      | #           return OBJECT_MAP[i]
      | #       end
      | #       i = i + 1
      | #   end
      | #   return OBJ_DEFAULT  # Return default pattern if not found
      | # end
      | 
      | def find_object_by_objectname(objectname):
      |     local i = 0
      |     #log_info("Trying to find object by color:", to_str(objectname))
      |     while (i < OBJECT_MAP.length()):
      |         if (OBJECT_MAP[i].obj_name == objectname):
      |             log_info("Object Model found: [" + to_str(OBJECT_MAP[i].description) + "]")
      |             return OBJECT_MAP[i]
      |         end
      |         i = i + 1
      |     end
      |     log_warning("no Object Model found for objectname:[" + to_str(objectname) + "]")
      |     return create_object()
      | end
      | 
      | def find_smallest_object():
      |     local i = 0
      |     local min_size = OBJECT_MAP[0].height
      |     #log_info("Trying to find object by color:", to_str(objectname))
      |     while (i < OBJECT_MAP.length()):
      |         if (OBJECT_MAP[i].height <= min_size and OBJECT_MAP[i].height != 0):
      |             log_info("smaller object found: [" + to_str(OBJECT_MAP[i].description) + "]")
      |             min_size = OBJECT_MAP[i].height
      |         end
      |         i = i + 1
      |     end
      |     return min_size
      | end
      | 
      | def find_gripper_config_by_objectname(objectname):
      | local i = 0
      | while (i < GRIPPER_CONFIG_MAP.length()):
      |     #log_info("gripper config:",to_str(GRIPPER_CONFIG_MAP[i]))
      |     if (GRIPPER_CONFIG_MAP[i].object == objectname):
      |         log_info("found gripper parameters [" + to_str(GRIPPER_CONFIG_MAP[i]) + "]")
      |         return GRIPPER_CONFIG_MAP[i]
      |     end
      |     i = i + 1
      | end
      | 
      | log_warning("no gripper parameters found for object type: " + to_str(objectname))
      | return create_gripper_config()
      | end
      | # Function to find a landmark by item
      | def find_landmark_by_id(lm_id):
      |     local i = 0
      |     while i < LANDMARK_MAP.length():
      |         if LANDMARK_MAP[i].lm_id == lm_id:
      |             log_info("found landmark with id(" + to_str(lm_id) + "): [" + to_str(LANDMARK_MAP[i].description) + "]")
      |             return LANDMARK_MAP[i]
      |         end
      |         i = i + 1
      |     end
      |     log_warning("landmark not found for lm_id [" + to_str(lm_id) + "]")
      |     return create_landmark()
      | end
      | # Function to find a landmark by item
      | def find_landmark_by_capture_pos(capture_pos):
      |     local i = 0
      |     while i < LANDMARK_MAP.length():
      |         if LANDMARK_MAP[i].capture_pos == capture_pos:
      |             log_info("found landmark by capture_pos [" + to_str(LANDMARK_MAP[i].description) + "]")
      |             return LANDMARK_MAP[i]
      |         end
      |         i = i + 1
      |     end
      |     log_warning("Landmark not found for capture_pos: [" + to_str(capture_pos) + "]")
      |     return create_landmark()
      | end
      | 
      | def update_landmark_by_capture_pos(capture_pos, lm_pos):
      |     local i = 0
      |     while i < LANDMARK_MAP.length():
      |         if LANDMARK_MAP[i].capture_pos == capture_pos:
      |             log_info("updated landmark from [" + to_str(LANDMARK_MAP[i].description) + "]")
      |             LANDMARK_MAP[i].actual_frame = lm_pos
      |             return True
      |         end
      |         i = i + 1
      |     end
      |     log_warning("Landmark not found for capture_pos: [" + to_str(capture_pos) + "]")
      |     return False
      | end
      | 
      | def update_landmark_by_id(lm_id,lm_pos):
      |     local i = 0
      |     while i < LANDMARK_MAP.length():
      |         if LANDMARK_MAP[i].lm_id == lm_id:
      |             log_info("updated landmark.actual_frame from [" + to_str(LANDMARK_MAP[i].description + "]"))
      |             LANDMARK_MAP[i].actual_frame = lm_pos
      |             return True
      |         end
      |         i = i + 1
      |     end
      |     log_warning("Landmark not found for lm_id " + to_str(lm_id))
      |     return False
      | end
      | 
      | def find_vision_config_by_frame(frame):
      |     local i = 0
      |     while i < VISION_CONFIG_MAP.length():
      |         if VISION_CONFIG_MAP[i].capture_pos == frame:
      |             log_info("Vision Config found: [" + to_str(VISION_CONFIG_MAP[i].description) + "]")
      |             return VISION_CONFIG_MAP[i]
      |         end
      |         i = i + 1
      |     end
      |     log_info("Vision Config not found for frame: " + to_str(frame))
      |     return create_vision_config()
      | end
      | 
      | def find_vision_config_by_itemid(id):
      |     local i = 0
      |     while i < VISION_CONFIG_MAP.length():
      |         if VISION_CONFIG_MAP[i].item_id == id:
      |             log_info("Vision Config found: [" + to_str(VISION_CONFIG_MAP[i].description) + "]")
      |             return VISION_CONFIG_MAP[i]
      |         end
      |         i = i + 1
      |     end
      |     log_info("Vision Config not found for item: " + to_str(id))
      |     return create_vision_config()
      | end
      | 
      | def find_inspect_config_by_itemid(id):
      |     local i = 0
      |     while i < INSPECT_CONFIG_MAP.length():
      |         if INSPECT_CONFIG_MAP[i].item_id == id:
      |             log_info("Inspect Config found: [" + to_str(INSPECT_CONFIG_MAP[i].description) + "]")
      |             return INSPECT_CONFIG_MAP[i]
      |         end
      |         i = i + 1
      |     end
      |     log_info("Inspect Config not found for item: " + to_str(id))
      |     return create_inspect_config()
      | end
    Script file /programs/04 Scripts/SCRIPT Device Robotiq Greifer v0.2.script
      | # ############ SCRIPT Device Robotiq Greifer ###############
      | # **********************************************************
      | # Customer          :   URG
      | # Product Name      :   uLabMobile
      | # **********************************************************
      | # Controller/Robot  :   UR5e
      | # Software          :   5.17
      | # Dependencies      :   Logs Script, Robotiq Gripper and Gripper Datastructure for args (Factory Script), URCAP Robotiq
      | # **********************************************************
      | # Author            :   D.Kreugel, P.Köhnke
      | # Copyright (c)     :   United Robotics Group Health and Food GmbH
      | #                       An der Riede 2
      | #                       28816 Stuhr
      | #                       Germany
      | # *********************************************************
      | # Description       :   Gripper Robotiq Device Interface for Robotiq E-Hand Gripper
      | # Version           :   0.2
      | # Created           :   18.07.2024
      | # Updated           :
      | # *********************************************************
      | # Modifications     :
      | #
      | # Date              :
      | # Name              :
      | # Reason            :
      | # *********************************************************
      | # TODO              :   documentation
      | 
      | # RobotiQ Gripper
      | ROBOTIQ_GRP_CLOSE = 0
      | ROBOTIQ_GRP_OPEN = 40
      | 
      | # #############FORCEMODE###############
      | ROBOTIQ_GRP_FORCE = struct(FULL=100, HALF=50, LOW=25, NONE=0)
      | 
      | # #############SPEED###################
      | ROBOTIQ_GRP_SPEED = struct(FAST=100, MEDIUM=50, SLOW=20)
      | 
      | # ############VALIDATION###############
      | ROBOTIQ_GRP_VALIDATION = struct(ON=1, OFF=0, SKIP=-1)
      | 
      | # struct(prepick=0, pick=0, place=0, force=0, speed=0, validation=0, object_type=0, description="default")
      | def gripper_robotiq_activate():
      |     return rq_activate_and_wait()
      | end
      | 
      | def gripper_robotiq_reset_and_activate():
      |     return rq_reset_and_activate()
      |     #return rq_reset()
      | end
      | 
      | def gripper_robotiq_is_activated():
      |     return rq_is_gripper_activated()
      | end
      | 
      | def gripper_robotiq_get_current_pos_mm():
      |     return rq_current_pos_mm()
      | end
      | # Function to check if the RobotiQ gripper has an object
      | def gripper_robotiq_has_object():
      |     result = rq_is_object_detected()
      |     if result == False:
      |         log_error("No object detected by the gripper")
      |     end
      |     return result
      | end
      | 
      | def gripper_robotiq_move_to_mm(mm):
      |     if(gripper_robotiq_is_activated() == False):
      |         gripper_robotiq_activate()
      |     end
      |     return rq_move_and_wait_mm(mm)
      | end
      | 
      | def gripper_robotiq_close():
      |     if(gripper_robotiq_is_activated() == False):
      |         gripper_robotiq_activate()
      |     end
      |     return rq_close_and_wait()
      | end
      | 
      | def gripper_robotiq_open():
      |     if(gripper_robotiq_is_activated() == False):
      |         gripper_robotiq_activate()
      |     end
      |     return rq_open_and_wait()
      | end
      | 
      | def gripper_robotiq_set_force(force):
      |     return rq_set_force_norm(force)
      | end
      | 
      | def gripper_robotiq_set_speed(velocity):
      |     return rq_set_speed_norm(velocity)
      | end
      | # Function to initialize the RobotiQ gripper
      | # args = struct(obj_type = object.obj_type, force = force, speed = speed, validation = validation, width = (prepick=2, pick=0, place=2))
      | def gripper_robotiq_init(args):
      |     log_info("args:"+to_str(args))
      |     gripper_robotiq_set_force(args.force)
      |     gripper_robotiq_set_speed(args.speed)
      |     if(gripper_robotiq_is_activated() == False):
      |         gripper_robotiq_activate()
      |     end
      |     log_info("Robotiq Gripper Initialized with arguments:" + to_str(args))
      |     return True
      | end
      | # Function to prepare the RobotiQ gripper for picking
      | # args = struct(obj_type = object.obj_type, force = force, speed = speed, validation = validation, width = (prepick=2, pick=0, place=2))
      | def gripper_robotiq_prepick(args):
      |     gripper_robotiq_init(args)
      | 
      |     if(args.width.prepick <= ROBOTIQ_GRP_CLOSE):
      |         rq_close_and_wait()
      |     elif(args.width.prepick >= ROBOTIQ_GRP_OPEN):
      |         rq_open_and_wait()
      |     else:
      |         rq_move_and_wait_mm(args.width.prepick)
      |     end
      | 
      |     log_info("Robotiq Gripper prepick with arguments:" + to_str(args))
      |     return True
      | end
      | 
      | # Function to place an object using the RobotiQ gripper
      | # args = struct(obj_type = object.obj_type, force = force, speed = speed, validation = validation, width = (prepick=2, pick=0, place=2))
      | def gripper_robotiq_place(args):
      |     gripper_robotiq_init(args)
      | 
      |     if(args.width.place <= ROBOTIQ_GRP_CLOSE):
      |         rq_close_and_wait()
      |     elif(args.width.place >= ROBOTIQ_GRP_OPEN):
      |         rq_open_and_wait()
      |     else:
      |         rq_move_and_wait_mm(args.width.place)
      |     end
      | 
      |     log_info("Gripper Place with arguments:"+ to_str(args))
      |     return True
      | end
      | 
      | # Function to pick an object using the RobotiQ gripper
      | # args = struct(obj_type = object.obj_type, force = force, speed = speed, validation = validation, width = (prepick=2, pick=0, place=2))
      | def gripper_robotiq_pick(args):
      |     gripper_robotiq_init(args)
      | 
      |     if(args.width.pick <= ROBOTIQ_GRP_CLOSE):
      |         rq_close_and_wait()
      |     elif(args.width.pick >= ROBOTIQ_GRP_OPEN):
      |         rq_open_and_wait()
      |     else:
      |         rq_move_and_wait_mm(args.width.pick)
      |     end
      | 
      |     log_info("Gripper Pick with arguments:" + to_str(args))
      | 
      |     if args.validation == ROBOTIQ_GRP_VALIDATION.ON:
      |         if gripper_robotiq_has_object() == False:
      |             log_error("Validation failed, no object detected")
      |             return False
      |         end
      |     end
      | 
      |     return True
      | end
      | 
      | 
      | # def gripper_robotiq_close_and_validate():
      | #     rq_close_and_wait()
      | #     if gripper_robotiq_has_object() == False:
      | #         log_error("Validation failed, no object detected")
      | #         return False
      | #     else:
      | #         return True
      | #     end
      | # end
    Script file /programs/04 Scripts/SCRIPT uLM Gripperconfig v0.6.script
      | ############# SCRIPT uLM Gripperconfig ###############
      | #*****************************************************
      | # Customer          :   URG
      | # Product Name      :   uLabMobile
      | #****************************************************
      | # Controller/Robot  :   UR5e
      | # Software          :   UR-Script
      | # Dependencies      :   physical Gripper and Datastructure from Factory for args -> Device Script and Implementations of the Functions
      | # How To            :   Assign all Functioncalls to the equivalent of the used Device Script
      | #****************************************************
      | # Author            :   D.Kreugel, P.Köhnke
      | # Copyright (c)     :   United Robotics Group Health and Food GmbH
      | #                       An der Riede 2
      | #                       28816 Stuhr
      | #                       Germany
      | #****************************************************
      | # Description       :   Defines all Gripperm related Parameters and Functions
      | # Version           :   0.6
      | # Created           :   18.07.2024
      | # Updated           :
      | #****************************************************
      | # Modifications     :   -> at the moment Gripperconfig linked to Robotiq Gripper Device Script
      | # Date              :   18.07.2017
      | # Name              :   D.Kreugel
      | # Reason            :   uLM Standard
      | #****************************************************
      | # TO DO             : Implement Activate and Reset Routine at the beginning or after an error depending on the state if an Object is gripped or not, documentation
      | 
      | 
      | 
      | # GRIPPER DEFINES
      | GRIPPER_CLOSE = ROBOTIQ_GRP_CLOSE
      | GRIPPER_OPEN = ROBOTIQ_GRP_OPEN
      | # #############FORCE###############
      | GRIPPER_FORCE = ROBOTIQ_GRP_FORCE
      | # #############SPEED###################
      | GRIPPER_SPEED = ROBOTIQ_GRP_SPEED
      | # ############VALIDATION###############
      | GRIPPER_VALIDATION = ROBOTIQ_GRP_VALIDATION
      | 
      | # takes force in %
      | def gripper_set_force(force):
      |     return gripper_robotiq_set_force(force)
      | end
      | 
      | # takes speed in %
      | def gripper_set_speed(velocity):
      |     return gripper_robotiq_set_speed(velocity)
      | end
      | 
      | def gripper_activate():
      |     return gripper_robotiq_activate()
      | end
      | 
      | def gripper_reset_and_activate():
      |     return gripper_robotiq_reset_and_activate()
      | end
      | 
      | def gripper_is_activated():
      |     return gripper_robotiq_is_activated()
      | end
      | 
      | def gripper_get_current_pos_mm():
      |     return gripper_robotiq_get_current_pos_mm()
      | end
      | 
      | def gripper_has_object():
      |     return gripper_robotiq_has_object()
      | end
      | 
      | def gripper_open():
      |     return gripper_robotiq_open()
      | end
      | 
      | def gripper_close():
      |     return gripper_robotiq_close()
      | end
      | 
      | def gripper_move_to_pos_mm(mm):
      |     return gripper_robotiq_move_to_mm(mm)
      | end
      | 
      | # args = struct(obj_type = object.obj_type, force = force, speed = speed, validation = validation, width = (prepick=2, pick=0, place=2))
      | def gripper_init(args):
      |     return gripper_robotiq_init(args)
      | end
      | 
      | # args = struct(obj_type = object.obj_type, force = force, speed = speed, validation = validation, width = (prepick=2, pick=0, place=2))
      | def gripper_prepick(args):
      |     return gripper_robotiq_prepick(args)
      | end
      | 
      | # args = struct(obj_type = object.obj_type, force = force, speed = speed, validation = validation, width = (prepick=2, pick=0, place=2))
      | def gripper_pick(args):
      |     return gripper_robotiq_pick(args)
      | end
      | 
      | # args = struct(obj_type = object.obj_type, force = force, speed = speed, validation = validation, width = (prepick=2, pick=0, place=2))
      | def gripper_place(args):
      |     return gripper_robotiq_place(args)
      | end
      | 
      | 
      | # def gripper_close_and_validate():
      | #     return gripper_robotiq_close_and_validate()
      | # end
    Script file /programs/04 Scripts/SCRIPT uLM Projectconfig 0.2.script
      | ############# SCRIPT uLM Projectconfig ###############
      | #*****************************************************
      | # Customer          :   URG
      | # Product Name      :   uLabMobile
      | #****************************************************
      | # Controller/Robot  :   UR5e
      | # Software          :   5.17
      | # Dependencies      :   Factory Script, Defines Script, relevant project knowledge about objects, patterns, items, commands, vision skills, landmarktypes and movements
      | # How To            :   Define Step by Step all Project Data by creating the objects and appending them to the assigned List, if you skip information
      | #                       the default value will be assigned -> give as many details as possible as the default values will not work in some cases
      | #****************************************************
      | # Author            :   D.Kreugel
      | # Copyright (c)     :   United Robotics Group Health and Food GmbH
      | #                       An der Riede 2
      | #                       28816 Stuhr
      | #                       Germany
      | #****************************************************
      | # Description       :   Project Related Configurations -> in the future will be configured by UGO
      | # Version           :   0.2
      | # Created           :   18.07.2024
      | # Updated           :
      | #****************************************************
      | # Modifications     :
      | # Date              :
      | # Name              :
      | # Reason            :
      | #****************************************************
      | # TO DO             :  Simplify Rack Assignment, create Enums for Choices that can be made and will be repeated in many projects, documentation
      | 
      | #
      | 
      | # Please Import DeviceScripts and Defines Script First as you may wanna use some of the Defined Variables here
      | 
      | # Define here the Objects that should be handled, add a new Object Type in the defines if necessary
      | # create_object(id=0, obj_name=0, height=0, width=0, color="default", material="default", description="default")
      | # struct(NONE=0, CC_SAMPLE=1, CC_RACK=2, COAG_SAMPLE=3, COAG_RACK=4, HEMA_SAMPLE=5, HEMA_RACK=6, INPUT_RACK=7, CF_RACK=8, ANY_SAMPLE=9, ANY_RACK=10)
      | #create_object(id=0, obj_name=0, height=0, width=0, obj_type = 0, description="default")
      | OBJECT_MAP.append(create_object(id=0, obj_name=Objects.NONE, obj_type=ObjectType.NONE, height=0, width=0, description="None Object"))
      | OBJECT_MAP.append(create_object(id=1, obj_name=Objects.CC_SAMPLE, obj_type=ObjectType.SAMPLE, height=108, width=15, description="BD Li-Heparin"))
      | OBJECT_MAP.append(create_object(id=2, obj_name=Objects.HEMA_SAMPLE, obj_type=ObjectType.SAMPLE, height=81, width=13, description="BD EDTA"))
      | OBJECT_MAP.append(create_object(id=3, obj_name=Objects.CC_SAMPLE, obj_type=ObjectType.SAMPLE, height=108, width=15, description="BD Li-Heparin"))
      | OBJECT_MAP.append(create_object(id=4, obj_name=Objects.HEMA_SAMPLE, obj_type=ObjectType.SAMPLE, height=81, width=13, description="Sarstedt EDTA"))
      | OBJECT_MAP.append(create_object(id=5, obj_name=Objects.CC_SAMPLE, obj_type=ObjectType.SAMPLE, height=110, width=15, description="Sarstedt Serum-Gel"))
      | OBJECT_MAP.append(create_object(id=6, obj_name=Objects.ANY_SAMPLE, obj_type=ObjectType.SAMPLE, height=110, width=15, description="Any Sample"))
      | OBJECT_MAP.append(create_object(id=7, obj_name=Objects.ANY_RACK, height=150, width=120, description="Any Rack"))
      | OBJECT_MAP.append(create_object(id=8, obj_name=Objects.CF_RACK, height=110, width=15, description="Centrifuge Rack"))
      | OBJECT_MAP.append(create_object(id=12, obj_name=Objects.COBAS_RACK, height=OBJECT_REFERENCE_HEIGHT, width=20, description="Cobas Rack"))
      | OBJECT_MAP.append(create_object(id=9, obj_name=Objects.TARA_SAMPLE, obj_type=ObjectType.SAMPLE, height=110, width=15, description="Tara Sample"))
      | OBJECT_MAP.append(create_object(id=10, obj_name=Objects.BUTTON, obj_type=ObjectType.BUTTON, height=0, width=0, description="Button"))
      | OBJECT_MAP.append(create_object(id=11, obj_name=Objects.XN550_DRAWER, height=OBJECT_REFERENCE_HEIGHT, width=25, description="XN550 Drawer"))
      | 
      | #create_sample(obj_id=0, diameter=0, color="", material="", description="")
      | SAMPLES = make_list(0,create_sample(),MAX_ITEM_OBJ)
      | SAMPLES.append(create_sample(obj_id=1, cap_diameter=17.4, raw_diameter=15.3, color="darkgreen", material="88", description="BD Li-Heparin -> decapped in Cobas"))
      | SAMPLES.append(create_sample(obj_id=1, cap_diameter=17.4, raw_diameter=15.3, color="darkgreen", material="80", description="BD Li-Heparin -> decapped in Cobas"))
      | SAMPLES.append(create_sample(obj_id=1, cap_diameter=17.4, raw_diameter=15.3, color="darkgreen", material="93", description="BD Li-Heparin -> decapped in archive"))
      | SAMPLES.append(create_sample(obj_id=2, cap_diameter=15.5, raw_diameter=12.3, color="violet", material="82", description="BD EDTA -> Sysmex ->Archive"))
      | SAMPLES.append(create_sample(obj_id=2, cap_diameter=15.5, raw_diameter=12.3, color="violet", material="91", description="BD EDTA ->Archive"))
      | SAMPLES.append(create_sample(obj_id=2, cap_diameter=15.5, raw_diameter=12.3, color="violet", material="96", description="BD EDTA ->Archive"))
      | SAMPLES.append(create_sample(obj_id=3, cap_diameter=17.4, raw_diameter=15.3, color="lightgreen", material="88", description="BD Li-Heparin -> decapped in Cobas"))
      | SAMPLES.append(create_sample(obj_id=3, cap_diameter=17.4, raw_diameter=15.3, color="lightgreen", material="93", description="BD Li-Heparin -> decapped in Archive"))
      | SAMPLES.append(create_sample(obj_id=3, cap_diameter=17.4, raw_diameter=15.3, color="lightgreen", material="97", description="BD Li-Heparin -> decapped in Archive"))
      | SAMPLES.append(create_sample(obj_id=4, cap_diameter=15.6, raw_diameter=12.3, color="red", material="82", description="BD EDTA -> Sysmex ->Archive"))
      | SAMPLES.append(create_sample(obj_id=4, cap_diameter=15.6, raw_diameter=12.3, color="red", material="91", description="BD EDTA -> Archive"))
      | SAMPLES.append(create_sample(obj_id=4, cap_diameter=15.6, raw_diameter=12.3, color="red", material="96", description="BD EDTA -> Archive"))
      | SAMPLES.append(create_sample(obj_id=5, cap_diameter=17.4, raw_diameter=15.3, color="brown", material="80", description="Sarstedt Serum-Gel -> decapped in Cobas"))
      | SAMPLES.append(create_sample(obj_id=5, cap_diameter=17.4, raw_diameter=15.3, color="brown", material="93", description="Sarstedt Serum-Gel -> decapped in Archive"))
      | 
      | # Gripper Configurations depending on the Object Type , add new force and speed in the Defines if necessary
      | # create_gripper_config(gripper_offset=struct(prepick=2, pick=0, place=2), force=0, speed=0, validation=0, object=create_object())
      | GRIPPER_CONFIG_MAP.append(create_gripper_config(gripper_offset=struct(prepick=2, pick=0, place=2), force=GRIPPER_FORCE.HALF, speed=GRIPPER_SPEED.MEDIUM, validation=GRIPPER_VALIDATION.ON, object=find_object_by_objectname(Objects.ANY_SAMPLE)))
      | GRIPPER_CONFIG_MAP.append(create_gripper_config(gripper_offset=struct(prepick=2, pick=0, place=2), force=GRIPPER_FORCE.FULL, speed=GRIPPER_SPEED.MEDIUM, validation=GRIPPER_VALIDATION.ON, object=find_object_by_objectname(Objects.ANY_RACK)))
      | GRIPPER_CONFIG_MAP.append(create_gripper_config(gripper_offset=struct(prepick=2, pick=0, place=2), force=GRIPPER_FORCE.HALF, speed=GRIPPER_SPEED.MEDIUM, validation=GRIPPER_VALIDATION.ON, object=find_object_by_objectname(Objects.CC_SAMPLE)))
      | GRIPPER_CONFIG_MAP.append(create_gripper_config(gripper_offset=struct(prepick=3, pick=0, place=3), force=GRIPPER_FORCE.HALF, speed=GRIPPER_SPEED.MEDIUM, validation=GRIPPER_VALIDATION.ON, object=find_object_by_objectname(Objects.HEMA_SAMPLE)))
      | GRIPPER_CONFIG_MAP.append(create_gripper_config(gripper_offset=struct(prepick=4, pick=0, place=4), force=GRIPPER_FORCE.HALF, speed=GRIPPER_SPEED.MEDIUM, validation=GRIPPER_VALIDATION.OFF, object=find_object_by_objectname(Objects.TARA_SAMPLE)))
      | GRIPPER_CONFIG_MAP.append(create_gripper_config(gripper_offset=struct(prepick=2, pick=0, place=2), force=GRIPPER_FORCE.FULL, speed=GRIPPER_SPEED.MEDIUM, validation=GRIPPER_VALIDATION.ON, object=find_object_by_objectname(Objects.CF_RACK)))
      | GRIPPER_CONFIG_MAP.append(create_gripper_config(gripper_offset=struct(prepick=2, pick=0, place=2), force=GRIPPER_FORCE.FULL, speed=GRIPPER_SPEED.MEDIUM, validation=GRIPPER_VALIDATION.ON, object=find_object_by_objectname(Objects.COBAS_RACK)))
      | GRIPPER_CONFIG_MAP.append(create_gripper_config(gripper_offset=struct(prepick=0, pick=0, place=0), force=GRIPPER_FORCE.HALF, speed=GRIPPER_SPEED.MEDIUM, validation=GRIPPER_VALIDATION.OFF, object=find_object_by_objectname(Objects.NONE)))
      | GRIPPER_CONFIG_MAP.append(create_gripper_config(gripper_offset=struct(prepick=0, pick=0, place=0), force=GRIPPER_FORCE.HALF, speed=GRIPPER_SPEED.MEDIUM, validation=GRIPPER_VALIDATION.OFF, object=find_object_by_objectname(Objects.BUTTON)))
      | GRIPPER_CONFIG_MAP.append(create_gripper_config(gripper_offset=struct(prepick=5, pick=25, place=5), force=GRIPPER_FORCE.HALF, speed=GRIPPER_SPEED.MEDIUM, validation=GRIPPER_VALIDATION.OFF, object=find_object_by_objectname(Objects.XN550_DRAWER)))
      | # create Patterns like Racks or Magazines
      | # easy if you define x and y regarding to the base coordinate system  if not you have to deal with transpose and or invert
      | # create_pattern(id=0, pattern_width=[0, 0], pattern_size=[0, 0], blocked=[-1, -1], obj_name=0, direction="X", transpose=False, invert=False, description="default")
      | # Objectss: NONE=0, CC_SAMPLE=1, CC_RACK=2, COAG_SAMPLE=3, COAG_RACK=4, HEMA_SAMPLE=5, HEMA_RACK=6, INPUT_RACK=7, CENTRIFUGE_RACK=8, ANY_SAMPLE=9, ANY_RACK=10
      | # ITEM_MODEL_MAP.append(create_pattern(id=0, pattern_width=[0, 0], pattern_size=[0, 0], blocked=[-1, -1, -1],  direction="X", transpose=False, invert=False, description="default"))
      | # ITEM_MODEL_MAP.append(create_pattern(id=1, pattern_width=[0.06, 0], pattern_size=[3, 1],  direction="X", description="Tara"))
      | # ITEM_MODEL_MAP.append(create_pattern(id=2, pattern_width=[0.183, 0.082], pattern_size=[10, 5], description="Sarstedt 50 D17 Rack"))
      | # ITEM_MODEL_MAP.append(create_pattern(id=3, pattern_width=[0.153, 0.067], pattern_size=[10, 5], description="Sarstedt 50 D13 Rack"))
      | # ITEM_MODEL_MAP.append(create_pattern(id=4, pattern_width=[0.06, 0.06], pattern_size=[3, 3], blocked=[5, -1, -1], description="Hettich Centrifuge Rack"))
      | # ITEM_MODEL_MAP.append(create_pattern(id=5, pattern_width=[0.093, 0.093], pattern_size=[2, 2],  description="Hettich Centrifuge Rack Magazin"))
      | # ITEM_MODEL_MAP.append(create_pattern(id=6, pattern_width=[0.08, 0.05], pattern_size=[5, 2], description="Sysmex XN 550 Rack"))
      | # ITEM_MODEL_MAP.append(create_pattern(id=7, pattern_width=[0.175, 0.078], pattern_size=[8, 4], description="URG Rack 40 D17"))
      | # ITEM_MODEL_MAP.append(create_pattern(id=8, pattern_width=[0.092, 0], pattern_size=[5, 1], description="Cobas Rack"))
      | # ITEM_MODEL_MAP.append(create_pattern(id=9, pattern_width=[0.245, 0.123], pattern_size=[3, 5], blocked=[9,11,12], description="Cobas Rack Magazin"))
      | # ITEM_MODEL_MAP.append(create_pattern(id=10, pattern_width=[0.237, 0.095], pattern_size=[11, 5], description="Atellica Rack 5x11"))
      | # ITEM_MODEL_MAP.append(create_pattern(id=11, pattern_width=[0.237, 0.095], pattern_size=[2, 2], description="Sensors LM"))
      | # ITEM_MODEL_MAP.append(create_pattern(id=12, pattern_width=[0.18, 0], pattern_size=[10, 1], description="Sysmex CS2500 Rack"))
      | # ITEM_MODEL_MAP.append(create_pattern(id=13, pattern_width=[0.310, 0.075], pattern_size=[13, 4], description="URG RACK 52 - Special Input"))
      | # ITEM_MODEL_MAP.append(create_pattern(id=14, pattern_width=[0.075, 0.075], pattern_size=[4, 6], description="URG RACK 24 - Special NoK"))
      | # ITEM_MODEL_MAP.append(create_pattern(id=15, pattern_width=[0.120, 0], pattern_size=[2, 1], description="XN550 Drawer"))
      | 
      | ITEM_MODEL_MAP.append(create_pattern(id=0, name="NONE", pattern_width=[0, 0], pattern_size=[0, 0], blocked=[-1, -1, -1],  direction="X", transpose=False, invert=False, description="default"))
      | ITEM_MODEL_MAP.append(create_pattern(id=1, name="TARA", pattern_width=[0.06, 0], pattern_size=[3, 1],  direction="X", description="Tara"))
      | ITEM_MODEL_MAP.append(create_pattern(id=4, name="CENTRIFUGE", pattern_width=[0.06, 0.06], pattern_size=[3, 3], blocked=[5, -1, -1], description="Hettich Centrifuge Rack"))
      | ITEM_MODEL_MAP.append(create_pattern(id=5, name="CENTRIFUGE_MAGAZINE", pattern_width=[0.093, 0.093], pattern_size=[2, 2],  description="Hettich Centrifuge Rack Magazin"))
      | ITEM_MODEL_MAP.append(create_pattern(id=6, name="SYSMEX_XN550", pattern_width=[0.08, 0.05], pattern_size=[5, 2], description="Sysmex XN 550 Rack"))
      | ITEM_MODEL_MAP.append(create_pattern(id=8, name="COBAS", pattern_width=[0.092, 0], pattern_size=[5, 1], description="Cobas Rack"))
      | ITEM_MODEL_MAP.append(create_pattern(id=9, name="COBAS_MAGAZINE", pattern_width=[0.245, 0.123], pattern_size=[3, 5], blocked=[9,11,12], description="Cobas Rack Magazin"))
      | ITEM_MODEL_MAP.append(create_pattern(id=13, name="INPUT", pattern_width=[0.310, 0.075], pattern_size=[13, 4], description="URG RACK 52 - Special Input"))
      | ITEM_MODEL_MAP.append(create_pattern(id=14, name="NOK", pattern_width=[0.075, 0.075], pattern_size=[4, 6], description="URG RACK 24 - Special NoK"))
      | ITEM_MODEL_MAP.append(create_pattern(id=15, name="DRAWER_XN550", pattern_width=[0.120, 0], pattern_size=[2, 1], description="XN550 Drawer"))
      | ITEM_MODEL_MAP.append(create_pattern(id=7, name="ARCHIVE", pattern_width=[0.175, 0.078], pattern_size=[8, 4], description="URG Rack 40 D17"))
      | 
      | 
      | 
      | 
      | 
      | 
      | # add a "skill" to the robots skillset the control system will send a string with the ls_item and action and here we will look if we have a matching skill to execute
      | # the item_modell defines the patterns which have to be used by the robot on multiple racks and or multiple samples in a rackpattern
      | # inner pattern is always dependung on the object that has to be moved and the outer pattern is the pattern for the containers where the objects are stored in.
      | # if racks have to be handled it is also an inner pattern cause the object to handle is the rack itself
      | # create_item(id=0, ls_item="default", frame=p[0,0,0,0,0,0], actionlist=create_action_list([]), item_model=create_item_model(), lm_id=0, description="default")
      | # create_item_model(inner=create_pattern(), outer=create_pattern(), description="default")
      | # ITEM_MAP.append(create_item(id=1, ls_item="Home", frame=F1_uLM_Home, actionlist=[ActionManipulator.MOVE_TO], description="uLM Move To Home"))
      | # ITEM_MAP.append(create_item(id=2, ls_item="InputStation", frame=F2_uLM_Input, actionlist=[ActionManipulator.PICK, ActionManipulator.PLACE], item_model=create_item_model(inner=Patterns.INPUT), description="uLM Pick and Place samples from Input"))
      | # ITEM_MAP.append(create_item(id=3, ls_item="InputCapture", frame=F3_Cap_Input, actionlist=[ActionCamera.INSPECT, ActionManipulator.MOVE_TO], description="uLM Inspect samples from Input and Move To Capture Position"))
      | # ITEM_MAP.append(create_item(id=4, ls_item="Bin", frame=F4_uLM_Bin, actionlist=[ActionManipulator.PLACE], description="uLM Place Cap to Bin"))
      | # ITEM_MAP.append(create_item(id=5, ls_item="StationaryGripper", frame=F5_uLM_Gripper, actionlist=[ActionManipulator.PICK, ActionManipulator.PLACE, ActionManipulator.DECAP, ActionManipulator.MOVE_TO, ActionManipulator.GRASP, ActionManipulator.RELEASE], description=" uLM stationary gripper"))
      | # ITEM_MAP.append(create_item(id=6, ls_item="CobasRack", frame=F6_uLM_Cobas_R, actionlist=[ActionManipulator.PICK, ActionManipulator.PLACE], item_model=create_item_model(outer=Patterns.COBAS_MAGAZINE), description="uLM Cobas Racks Pick and Place"))
      | # ITEM_MAP.append(create_item(id=7, ls_item="CobasMagazine", frame=F7_uLM_Coba_Mag, actionlist=[ActionManipulator.PICK, ActionManipulator.PLACE], item_model=create_item_model(inner=Patterns.COBAS, outer=Patterns.COBAS_MAGAZINE), description="uLM Cobas Magazine Samples Pick and Place"))
      | # ITEM_MAP.append(create_item(id=8, ls_item="DetectCobasRacks", frame=F8_Cap_Cobas_LM, actionlist=[ActionCamera.DETECT_OBJECTS, ActionManipulator.MOVE_TO], lm_id=2, description="uLM Cobas Rack Detection and Move To Capture"))
      | # ITEM_MAP.append(create_item(id=9, ls_item="TaraMagazine", frame=F9_uLM_Tara, actionlist=[ActionManipulator.PICK, ActionManipulator.PLACE], item_model=create_item_model(inner=Patterns.TARA), description="uLM Centrifuge Tara Pick and Place"))
      | # ITEM_MAP.append(create_item(id=10, ls_item="CentrifugeCapture", frame=F10_Cap_CF, actionlist=[ActionManipulator.MOVE_TO, ActionCamera.DETECT], lm_id=1, description="Centrifuge Device Move to Capture Pos and Detect Landmarks"))
      | # ITEM_MAP.append(create_item(id=11, ls_item="Centrifuge", frame=F11_CF_PiPl, actionlist=[ActionManipulator.PICK, ActionManipulator.PLACE], description="Centrifuge Device Rack Pick and Place"))
      | # ITEM_MAP.append(create_item(id=12, ls_item="CentrifugeMagazine", frame=F12_uLM_CF_Mag, actionlist=[ActionManipulator.PICK, ActionManipulator.PLACE], item_model=create_item_model(inner=Patterns.CENTRIFUGE, outer=Patterns.CENTRIFUGE_MAGAZINE), description=" uLM Centrifuge Magazin Pick and Place"))
      | # ITEM_MAP.append(create_item(id=13, ls_item="CentrifugeRack", frame=F13_uLM_CF_R, actionlist=[ActionManipulator.PICK, ActionManipulator.PLACE], item_model=create_item_model(outer=Patterns.CENTRIFUGE_MAGAZINE), description="uLM Centrifuge Magazin Pick and Place Racks"))
      | # ITEM_MAP.append(create_item(id=14, ls_item="DailyArchive", frame=F14_uLM_Archive, actionlist=[ActionManipulator.PICK, ActionManipulator.PLACE], item_model=create_item_model(inner=Patterns.ARCHIVE), description="uLM Pick and Place samples from Archive Rack"))
      | # ITEM_MAP.append(create_item(id=15, ls_item="NokRack", frame=F15_uLM_Nok, actionlist=[ActionManipulator.PICK, ActionManipulator.PLACE], item_model=create_item_model(inner=Patterns.NOK), description="uLM Pick and Place samples from Nok Rack"))
      | # ITEM_MAP.append(create_item(id=16, ls_item="CobasInput", frame=F16_Cobas_Input, actionlist=[ActionManipulator.PLACE], description="uLM Place Cobasrack in Cobas Device"))
      | # ITEM_MAP.append(create_item(id=17, ls_item="CobasInputCapture", frame=F17_Cobas_Cap, actionlist=[ActionCamera.DETECT, ActionManipulator.MOVE_TO], lm_id=3, description="uLM Place Cobasrack in Cobas Device"))
      | # ITEM_MAP.append(create_item(id=18, ls_item="XN550Input", frame=F18_XN550_Input, actionlist=[ActionManipulator.PICK, ActionManipulator.PLACE], item_model=create_item_model(inner=Patterns.SYSMEX_XN550, outer=Patterns.DRAWER_XN550), lm_id=4, description="uLM Pick and Place Samples in or out of XN550 Racks"))
      | # ITEM_MAP.append(create_item(id=19, ls_item="XN550Capture", frame=F19_XN550_Cap, actionlist=[ActionCamera.DETECT, ActionManipulator.MOVE_TO], lm_id=4, description="uLM Move To and Capture LM XN550"))
      | # ITEM_MAP.append(create_item(id=20, ls_item="XN550Drawer", frame=F20_XN550_Draw, actionlist=[ActionManipulator.DRAWER_OPEN, ActionManipulator.DRAWER_CLOSE], item_model=create_item_model(inner=Patterns.DRAWER_XN550), lm_id=4, description="uLM Open and close Drawer XN550"))
      | # ITEM_MAP.append(create_item(id=21, ls_item="XN550Button", frame=F21_XN550_Btn, actionlist=[ActionManipulator.PUSH], lm_id=4, description="uLM Push XN550 Button"))
      | # ITEM_MAP.append(create_item(id=22, ls_item="AMR", frame=p[0,0,0,0,0,0], actionlist=[ActionAMR.READ, ActionAMR.LOAD_MISSION, ActionAMR.START_MISSION, ActionAMR.NAVIGATE, ActionAMR.ACKNOWLEDGE], description="all AMR actions"))
      | 
      | 
      | 
      | # ITEM_MAP.append(create_item(id=31, ls_item="TestLM", frame=TestLM, actionlist=[ActionManipulator.PICK, ActionManipulator.PLACE], item_model=create_item_model(inner=Rack.SYSMEX_CS2500), lm_id=5, description="LM Test"))
      | # Fills the Vision Config List with Projectrelated Data
      | # workspaceid and skillid are highly robominds related so probably will not stay like this in the future
      | # sample detection: dx and dy are used to calculate the positions in a rack and given by the offset which will be applied in order to assign the sample to a place in the rack
      | # create_vision_config(workspace_id="", skill_id="", item_id=-1, capture_pos=p[0,0,0,0,0,0], dx=0, dy=0, target_origin=p[0,0,0,0,0,0], selector="default", description="default")
      | # VISION_CONFIG_MAP.append(create_vision_config(workspace_id="96017791-f581-4e9e-93da-6951695fccc8", skill_id="8885cfe1-6784-4293-bd26-52ebdc67bf95", capture_pos=F10_Cap_CF, target_origin=p[0,0,0,0,0,0], item_id=11, description="LM Detect CF"))
      | # VISION_CONFIG_MAP.append(create_vision_config(workspace_id="96017791-f581-4e9e-93da-6951695fccc8", skill_id="8885cfe1-6784-4293-bd26-52ebdc67bf95", capture_pos=F8_Cap_Cobas_LM, target_origin=p[0,0,0,0,0,0], item_id=8, description="LM Detect Cobas Racks"))
      | # VISION_CONFIG_MAP.append(create_vision_config(workspace_id="8f0ad01c-dc36-4fdd-b295-0b6b4a38b89a", skill_id="afdc9e13-ea83-40d6-a805-bb041453d2e5", capture_pos=F3_Cap_Input, target_origin=F2_uLM_Input, item_id=3, description="Lab Solution Input Capture"))
      | # VISION_CONFIG_MAP.append(create_vision_config(workspace_id="96017791-f581-4e9e-93da-6951695fccc8", skill_id="8885cfe1-6784-4293-bd26-52ebdc67bf95", capture_pos=F19_XN550_Cap, target_origin=F18_XN550_Input, item_id=18, description="Input XN550"))
      | # VISION_CONFIG_MAP.append(create_vision_config(workspace_id="96017791-f581-4e9e-93da-6951695fccc8", skill_id="8885cfe1-6784-4293-bd26-52ebdc67bf95", capture_pos=F19_XN550_Cap, target_origin=POS_Z, item_id=19, description="LM Detect XN550F"))
      | # VISION_CONFIG_MAP.append(create_vision_config(workspace_id="96017791-f581-4e9e-93da-6951695fccc8", skill_id="8885cfe1-6784-4293-bd26-52ebdc67bf95", capture_pos=F10_Cap_CF, target_origin=POS_Z, item_id=10, description="LM Detect CF"))
      | # VISION_CONFIG_MAP.append(create_vision_config(workspace_id="96017791-f581-4e9e-93da-6951695fccc8", skill_id="8885cfe1-6784-4293-bd26-52ebdc67bf95", capture_pos=F19_XN550_Cap, target_origin=F20_XN550_Draw, item_id=20, description="Drawer XN550"))
      | # VISION_CONFIG_MAP.append(create_vision_config(workspace_id="96017791-f581-4e9e-93da-6951695fccc8", skill_id="8885cfe1-6784-4293-bd26-52ebdc67bf95", capture_pos=F19_XN550_Cap, target_origin=F21_XN550_Btn, item_id=21, description="Button XN550"))
      | # VISION_CONFIG_MAP.append(create_vision_config(workspace_id="96017791-f581-4e9e-93da-6951695fccc8", skill_id="8885cfe1-6784-4293-bd26-52ebdc67bf95", capture_pos=TestLMCap, target_origin=p[0,0,0,0,0,0], item_id=30, description="Button XN550"))
      | # VISION_CONFIG_MAP.append(create_vision_config(workspace_id="96017791-f581-4e9e-93da-6951695fccc8", skill_id="8885cfe1-6784-4293-bd26-52ebdc67bf95", capture_pos=TestLMCap, target_origin=TestLM, item_id=31, description="Button XN550"))
      | 
      | # VISION_CONFIG_MAP.append(create_vision_config(workspace_id="96017791-f581-4e9e-93da-6951695fccc8", skill_id="8885cfe1-6784-4293-bd26-52ebdc67bf95", target_origin=p[0,0,0,0,0,0], item_id=11, description="LM Detect CF"))
      | # VISION_CONFIG_MAP.append(create_vision_config(workspace_id="96017791-f581-4e9e-93da-6951695fccc8", skill_id="8885cfe1-6784-4293-bd26-52ebdc67bf95", target_origin=p[0,0,0,0,0,0], item_id=8, description="LM Detect Cobas Racks"))
      | # VISION_CONFIG_MAP.append(create_vision_config(workspace_id="8f0ad01c-dc36-4fdd-b295-0b6b4a38b89a", skill_id="afdc9e13-ea83-40d6-a805-bb041453d2e5", target_origin=F2_uLM_Input, item_id=3, description="Lab Solution Input Capture"))
      | # VISION_CONFIG_MAP.append(create_vision_config(workspace_id="96017791-f581-4e9e-93da-6951695fccc8", skill_id="8885cfe1-6784-4293-bd26-52ebdc67bf95", target_origin=F18_XN550_Input, item_id=18, description="Input XN550"))
      | # VISION_CONFIG_MAP.append(create_vision_config(workspace_id="96017791-f581-4e9e-93da-6951695fccc8", skill_id="8885cfe1-6784-4293-bd26-52ebdc67bf95", target_origin=POS_Z, item_id=19, description="LM Detect XN550F"))
      | # VISION_CONFIG_MAP.append(create_vision_config(workspace_id="96017791-f581-4e9e-93da-6951695fccc8", skill_id="8885cfe1-6784-4293-bd26-52ebdc67bf95", target_origin=POS_Z, item_id=10, description="LM Detect CF"))
      | # VISION_CONFIG_MAP.append(create_vision_config(workspace_id="96017791-f581-4e9e-93da-6951695fccc8", skill_id="8885cfe1-6784-4293-bd26-52ebdc67bf95", target_origin=F20_XN550_Draw, item_id=20, description="Drawer XN550"))
      | # VISION_CONFIG_MAP.append(create_vision_config(workspace_id="96017791-f581-4e9e-93da-6951695fccc8", skill_id="8885cfe1-6784-4293-bd26-52ebdc67bf95", target_origin=F21_XN550_Btn, item_id=21, description="Button XN550"))
      | # VISION_CONFIG_MAP.append(create_vision_config(workspace_id="96017791-f581-4e9e-93da-6951695fccc8", skill_id="8885cfe1-6784-4293-bd26-52ebdc67bf95", target_origin=p[0,0,0,0,0,0], item_id=30, description="Button XN550"))
      | # VISION_CONFIG_MAP.append(create_vision_config(workspace_id="96017791-f581-4e9e-93da-6951695fccc8", skill_id="8885cfe1-6784-4293-bd26-52ebdc67bf95", target_origin=TestLM, item_id=31, description="Button XN550"))
      | 
      | # local inputrack = find_pattern_by_name("INPUT")
      | # INSPECT_CONFIG_MAP.append(create_inspect_config(item_id=3, dx=inputrack.pattern_width[0]/(inputrack.pattern_size[0]-1), dy=inputrack.pattern_width[1]/(inputrack.pattern_size[1]-1), rack_size=inputrack.pattern_size , description="Input Capture"))
      | # # Fills the Landmark List with Projectrelated Data
      | # # create_landmark(lm_id=0, marker_id=-1, marker_size=0.1, marker_type="aruco_7x7", capture_pos=p[0,0,0,0,0,0], init_frame=p[0,0,0,0,0,0], search_offset=[0,0,0], actual_frame=p[0,0,0,0,0,0], description="")
      | # LANDMARK_MAP.append(create_landmark(lm_id=1, marker_id=3, marker_size=0.1, marker_type="aruco_7x7", capture_pos = F10_Cap_CF, init_frame=p[-0.617789, -0.065471, 0.07918, 0.020983, -0.012695, 1.512066], search_offset=[0.15, 0.15, 0.1], actual_frame=p[-0.617789, -0.065471, 0.07918, 0.020983, -0.012695, 1.512066], description="LM CF Lid"))
      | # LANDMARK_MAP.append(create_landmark(lm_id=2, marker_id=-1, marker_size=0.0085, marker_type="aruco_4x4", capture_pos = F8_Cap_Cobas_LM, init_frame=p[0,0,0,0,0,0], search_offset=[0.15, 0.15, 0.1], actual_frame=POS_Z, description="LM Cobas Rack Detection"))
      | # LANDMARK_MAP.append(create_landmark(lm_id=3, marker_id=0, marker_size=0.1, marker_type="aruco_7x7", capture_pos = F17_Cobas_Cap, init_frame=p[-0.667,-0.194,0.100,0,0,0], search_offset=[0.15, 0.15, 0.1], actual_frame=POS_Z, description="LM Cobas Cap"))
      | # LANDMARK_MAP.append(create_landmark(lm_id=4, marker_id=4, marker_size=0.1, marker_type="aruco_7x7", capture_pos = F19_XN550_Cap, init_frame=p[0.124,-0.976,0.355,-0.008,0.025,3.131], search_offset=[0.15, 0.15, 0.1], actual_frame=p[0,0,0,0,0,0], description="LM XN550 Cap"))
      | # LANDMARK_MAP.append(create_landmark(lm_id=5, marker_id=0, marker_size=0.1, marker_type="aruco_7x7", capture_pos = TestLMCap, init_frame=p[-0.49,-0.144,0.092,0,-0.008,0.001], search_offset=[0.15, 0.15, 0.1], actual_frame=POS_Z, description="LM Test"))
      | # # Configuration of all movement related parameters
      | # # create_movement(id=0, hh_approach=POS_Z, h_approach=POS_Z, approach=POS_Z, h_target=POS_Z, target=POS_Z, retract=POS_Z, h_retract=POS_Z, hh_retract=POS_Z, h_frame=POS_Z, frame=POS_Z, speed=1, acceleration=1, description="default")
      | # MOVEMENT_MAP.append(create_movement(description="TestLMCap", frame=TestLMCap, actionlist=[ActionManipulator.MOVE_TO]))
      | # MOVEMENT_MAP.append(create_movement(description="TestLM", frame=TestLM, actionlist=[ActionManipulator.PICK,ActionManipulator.PLACE],
      | #         approach=p[0,0,0.1,0,0,0],
      | #         retract=p[0,0,0.1,0,0,0]))
      | # MOVEMENT_MAP.append(create_movement(description="Home - MOVE_TO", frame=F1_uLM_Home, actionlist=[ActionManipulator.MOVE_TO]))
      | # MOVEMENT_MAP.append(create_movement(description="Input - PICK&PLACE", frame=F2_uLM_Input, actionlist=[ActionManipulator.PICK,ActionManipulator.PLACE],
      | #         approach=p[0,0,0.1,0,0,0],
      | #         retract=p[0,0,0.1,0,0,0]))
      | # MOVEMENT_MAP.append(create_movement(description="Capture Input - MOVE_TO", frame=F3_Cap_Input, actionlist=[ActionManipulator.MOVE_TO]))
      | # MOVEMENT_MAP.append(create_movement(description="BIN - PLACE", frame=F4_uLM_Bin, actionlist=[ActionManipulator.PLACE],
      | #         approach=p[0,0,0.1,0,0,0],
      | #         retract=p[0,0,0.1,0,0,0]))
      | # MOVEMENT_MAP.append(create_movement(description="Gripper - Move To", frame=F5_uLM_Gripper, actionlist=[ActionManipulator.MOVE_TO],
      | #         approach=p[0,0,0.1,0,0,0]))
      | # MOVEMENT_MAP.append(create_movement(description="Gripper - Pick", frame=F5_uLM_Gripper, actionlist=[ActionManipulator.PICK],
      | #         retract=p[0,0,0.1,0,0,0]))
      | # MOVEMENT_MAP.append(create_movement(description="Gripper - Place", frame=F5_uLM_Gripper, actionlist=[ActionManipulator.PLACE],
      | #         approach=p[0,0,0.1,0,0,0]))
      | # MOVEMENT_MAP.append(create_movement(description="CobasRack Pick & Place", frame=F6_uLM_Cobas_R, actionlist=[ActionManipulator.PICK,ActionManipulator.PLACE],
      | #         approach=p[0,0,0.1,0,0,0],
      | #         target=p[0,0,0,0,0,d2r(90)],
      | #         retract=p[0,0,0.1,0,0,0]))
      | # MOVEMENT_MAP.append(create_movement(description="CobasMagazine Pick & Place", frame=F7_uLM_Coba_Mag, actionlist=[ActionManipulator.PICK,ActionManipulator.PLACE],
      | #         approach=p[0,0,0.1,0,0,0],
      | #         target=p[0,0,0,0,0,-d2r(90)],
      | #         retract=p[0,0,0.1,0,0,0]))
      | # MOVEMENT_MAP.append(create_movement(description="Capture Position Cobas Landmarks", frame=F8_Cap_Cobas_LM, actionlist=[ActionManipulator.MOVE_TO]))
      | # MOVEMENT_MAP.append(create_movement(description="TaraMagazine - PICK & PLACE", frame=F9_uLM_Tara, actionlist=[ActionManipulator.PICK,ActionManipulator.PLACE],
      | #         approach=p[0,0,0.13,0,0,0],
      | #         target=p[0,0,0,0,0,-d2r(90)],
      | #         retract=p[0,0,0.13,0,0,0]))
      | # MOVEMENT_MAP.append(create_movement(description="Capture Position - Centrifuge LM", frame=F10_Cap_CF,actionlist=[ActionManipulator.MOVE_TO]))
      | # MOVEMENT_MAP.append(create_movement(description="Pick and Place Racks - Centrifuge Lid", frame=F11_CF_PiPl, actionlist=[ActionManipulator.PICK,ActionManipulator.PLACE],
      | #         approach=p[0,0,0.3,0,0,0],
      | #         retract=p[0,0,0.3,0,0,0]))
      | # MOVEMENT_MAP.append(create_movement(description="Pick and Place Samples - Centrifuge on uLM", frame=F12_uLM_CF_Mag, actionlist=[ActionManipulator.PICK,ActionManipulator.PLACE],
      | #         approach=p[0,0,0.13,0,0,0],
      | #         retract=p[0,0,0.13,0,0,0]
      | #         ))
      | # MOVEMENT_MAP.append(create_movement(description="Pick and Place Racks - Centrifuge on uLM", frame=F13_uLM_CF_R, actionlist=[ActionManipulator.PICK,ActionManipulator.PLACE],
      | #         approach=p[0,0,0.15,0,0,0],
      | #         retract=p[0,0,0.15,0,0,0]
      | #         ))
      | 
      | # MOVEMENT_MAP.append(create_movement(description="Pick and Place Samples XN550 Racks in Device", frame=F18_XN550_Input, actionlist=[ActionManipulator.PICK,ActionManipulator.PLACE],
      | #         approach=p[0,0,0.1,0,0,0],
      | #         target = p[0,0,0,0,0,d2r(90)],
      | #         retract=p[0,0,0.1,0,0,0]
      | #         ))
      | # MOVEMENT_MAP.append(create_movement(description="Capture LM XN550", frame=F19_XN550_Cap, actionlist=[ActionManipulator.MOVE_TO]))
      | # MOVEMENT_MAP.append(create_movement(description="Open XN550 Drawer ", frame=F20_XN550_Draw, actionlist=[ActionManipulator.DRAWER_OPEN],
      | #         h_approach=p[0.07,0,0.1,0,0,0],
      | #         approach=p[0,0,0.1,0,0,0],
      | #         target = p[0,0,0,0,0,d2r(90)],
      | #         retract=p[0.07,0,0,0,0,0],
      | #         h_retract=p[0.07,0,0.1,0,0,0]
      | #         ))
      | # MOVEMENT_MAP.append(create_movement(description="Close XN550 Drawer ", frame=F20_XN550_Draw, actionlist=[ActionManipulator.DRAWER_CLOSE],
      | #         h_approach=p[0.07,0,0.1,0,0,0],
      | #         approach=p[0.07,0,0,0,0,0],
      | #         target = p[0,0,0,0,0,d2r(90)],
      | #         retract=p[0,0,0.1,0,0,0],
      | #         h_retract=p[0.07,0,0.1,0,0,0]
      | #         ))
      | # MOVEMENT_MAP.append(create_movement(description="Push XN550 Button ", frame=F21_XN550_Btn, actionlist=[ActionManipulator.PUSH],
      | #         approach=p[0,0,0.15,0,0,0],
      | #         retract=p[0,0,0.15,0,0,0]
      | #         ))
      | # MOVEMENT_MAP.append(create_movement(description="Capture Position 2 Input", frame=F_Cap_Input2,actionlist=[ActionManipulator.MOVE_TO]))
    Script file /programs/04 Scripts/SCRIPT Objects V0.1.script
      | #*****************************************************
      | # customer          :   INTERNAL
      | # project name      :
      | #****************************************************
      | # controller        :   UR
      | # software          :   5.17.3
      | #****************************************************
      | # author            :   P. Koehnke
      | # Copyright (c)     :   United Robotics Group
      | #                       An der Riede 2
      | #                       28816 Stuhr
      | #                       Germany
      | #****************************************************
      | # description       :   object database
      | # version:      	:   0.1
      | # created           :   09.10.2024
      | # updated           :
      | #****************************************************
      | # modifications     :
      | #
      | # date              :
      | # name              :
      | # reason            :
      | #****************************************************
      | 
      | def create_object_2(id=0, name="", type=0, dimension=struct(length=0, width=0, height=0, diameter=0), gripper_offset=p[0,0,0,0,0,0]):
      |     return struct(id=id, name=name, type=type, dimension=dimension, gripper_offset=gripper_offset)
      | end
      | 
      | OBJ = create_object_2()
      | OBJs = make_list(0, create_object_2(), 50)
      | 
      | OBJs.append(create_object_2(id=1, name="rack centrifuge", type=1, dimension=struct(length=0, width=0, height=0.106, diameter=0.020), gripper_offset=p[0,0,0.095,0,0,2.356]))
      | OBJs.append(create_object_2(id=2, name="sample tube 1", type=2, dimension=struct(length=0, width=0, height=0.106, diameter=0.015), gripper_offset=p[0,0,0,0,0,0]))
      | OBJs.append(create_object_2(id=3, name="rack sarstedt", type=3, dimension=struct(length=0, width=0, height=0.100, diameter=0.020), gripper_offset=p[0,0,0,0,0,0]))
      | OBJs.append(create_object_2(id=4, name="Lab bottle", type=4, dimension=struct(length=0, width=0, height=0.100, diameter=0.030), gripper_offset=p[0,0,0.2,0,0,0]))
      | OBJs.append(create_object_2(id=5, name="Vial", type=5, dimension=struct(length=0, width=0, height=0.100, diameter=0.0275), gripper_offset=p[0,0,0,0,0,0]))
      | OBJs.append(create_object_2(id=6, name="Container", type=6, dimension=struct(length=0.0, width=0.0, height=0, diameter=0.0), gripper_offset=p[0,0,0,0,0,0]))
      | OBJs.append(create_object_2(id=7, name="Target_container", type=7, dimension=struct(length=0.06, width=0.06, height=0.134, diameter=0.05), gripper_offset=p[0,0,0,0,0,0]))
      | OBJs.append(create_object_2(id=8, name="Spatula", type=8, dimension=struct(length=0.03, width=0.03, height=0.23, diameter=0.05), gripper_offset=p[0,0,0,0,0,0]))
      | OBJs.append(create_object_2(id=9, name="rack pipet", type=9, dimension=struct(length=0.03, width=0.03, height=0.23, diameter=0.05), gripper_offset=p[0,0,0,0,0,0]))
      | 
      | def create_jig_2(id=0, name="", type=0, capacity=0, jig_offset=p[0,0,0,0,0,0]):
      |     # iformation about used jigs
      |     return struct(id=id, name=name, type=type, capacity=capacity, jig_offset=jig_offset)
      | end
      | 
      | JIG2 = create_jig_2()
      | JIGs = make_list(0, create_jig_2(), 20)
      | 
      | JIGs.append(create_jig_2(id=1, name="3FG", type=1, capacity=1, jig_offset=p[0,0,0,0,0,0]))
      | JIGs.append(create_jig_2(id=2, name="jig input", type=2, capacity=1, jig_offset=p[0,0,0,0,0,-3.927]))
      | JIGs.append(create_jig_2(id=3, name="jig output", type=3, capacity=1, jig_offset=p[0,0,0,0,0,0.78]))
      | JIGs.append(create_jig_2(id=6, name="jig bin", type=6, capacity=1, jig_offset=p[0,0,0,0,0,0]))
      | JIGs.append(create_jig_2(id=7, name="jig sarstedt racks", type=7, capacity=1, jig_offset=p[0,0,-0.02,0,0,0]))
      | JIGs.append(create_jig_2(id=8, name="NoK Bin", type=8, capacity=1, jig_offset=p[0,0,0,0,0,0]))
      | JIGs.append(create_jig_2(id=9, name="Pick bott jig", type=9, capacity=1, jig_offset=p[0,0,0,0,0,0]))
      | JIGs.append(create_jig_2(id=10, name="Place bott jig", type=10, capacity=1, jig_offset=p[0,0,0,0,0,0]))
      | JIGs.append(create_jig_2(id=11, name="bottle shake jig", type=11, capacity=1, jig_offset=p[0,0,0,0,0,0]))
      | JIGs.append(create_jig_2(id=12, name="Pick Vial jig", type=12, capacity=1, jig_offset=p[0,0,0,0,0,0]))
      | JIGs.append(create_jig_2(id=13, name="Place Vial jig", type=13, capacity=1, jig_offset=p[0,0,0,0,0,0]))
      | JIGs.append(create_jig_2(id=14, name="Liquid transfer jig", type=14, capacity=1, jig_offset=p[0,0,0,0,0,0]))
      | JIGs.append(create_jig_2(id=15, name="Pick station jig", type=15, capacity=1, jig_offset=p[0,0,0,0,0,0]))
      | JIGs.append(create_jig_2(id=16, name="Place station jig", type=16, capacity=1, jig_offset=p[0,0,0,0,0,0]))
      | JIGs.append(create_jig_2(id=17, name="Weigh station jig", type=17, capacity=1, jig_offset=p[0,0,0,0,0,0]))
      | JIGs.append(create_jig_2(id=18, name="Pick station 1", type=18, capacity=1, jig_offset=p[0,0,0,0,0,0]))
      | JIGs.append(create_jig_2(id=19, name="Pick station 2", type=19, capacity=1, jig_offset=p[0,0,0,0,0,0]))
      | JIGs.append(create_jig_2(id=20, name="Pick station 3", type=20, capacity=1, jig_offset=p[0,0,0,0,0,0]))
      | JIGs.append(create_jig_2(id=21, name="Tilt station jig", type=21, capacity=1, jig_offset=p[0,0,0,0,0,0]))
    Script file /programs/04 Scripts/Powder_all copy.script
      | #global SERVER_IP   = "192.168.12.139"
      | 
      | 
      | global tcp_dosing = p[0,0,0.15052,3.1415,0,0]
      | global tcp_default = p[0,0,0.161,3.1415,0,0]
      | 
      | global container_id = 0
      | global powder_id  = 0
      | global bulk_density = 0
      | global H          = 0
      | global H_c          = 0
      | global mouth_d     = 0
      | global mouth_sh    = 0
      | global length_c     = 0
      | global diameter   = 0
      | global empty_weight_g  = 0
      | global volume_ml    = 0
      | global shape_code   = 0
      | global flow_code   = 0
      | global shape = ""
      | global Flowability = ""
      | global full_weight_g = 0
      | global cent_edge = 0
      | global pick_2_base = 0.2 # distance from tcp to base of picking table
      | global wall_thickness = 0.002
      | 
      | def read_db_data():
      | 
      |   socket_open(SERVER_IP, SERVER_PORT)
      |   sleep(0.5)
      |   socket_send_string("GET_DATACODE_FLOATS")
      |   sleep(5)
      | 
      |   local fl = socket_read_ascii_float(14)
      |   socket_close()
      | 
      |   global container_id = fl[1]
      |   global powder_id = fl[2]
      |   global bulk_density = fl[3]
      |   global H          = fl[4]/1000
      |   global H_c          = fl[5]/1000
      |   global mouth_d     = fl[6]/1000
      |   global mouth_sh    = fl[7]/1000
      |   global length_c     = fl[8]/1000
      |   global diameter   = fl[9]/1000
      |   global empty_weight_g = fl[10]
      |   global volume_ml    = fl[11]
      |   global full_weight_g = fl[12]
      |   global flow_code   = fl[13]
      |   global shape_code   = fl[14]
      | 
      | 	if (flow_code == 1.0):
      | 	  global Flowability = "MEDIUM"
      | 	elif (flow_code == 2.0):
      | 	  global Flowability = "LOW"
      | 	else:
      | 	  global Flowability = "HIGH"
      | 	end
      | 
      |   if ( shape_code == 1.0):
      | 	shape = "cylindrical"
      | 	cent_edge =  diameter
      |   else:
      | 	shape = "cubical"
      | 	cent_edge =  length_c
      |   end
      | 
      | end
      | 
      | def send_picking_info(Pow_name, target_weight):
      |   socket_open(SERVER_IP, SERVER_PORT)
      |   cmd = "PICK:"+Pow_name+";"+to_str(target_weight)
      |   socket_send_string(cmd)
      |   sleep(0.1)
      |   socket_close()
      | end
      | 
      | #### POTS ####
      | def tilt_send(angle):
      | 	socket_open(SERVER_IP, SERVER_PORT)
      | 	angle = 92.0 - angle
      | 	socket_send_string("TILT:"+to_str(angle))
      | 	sync()
      | 	sleep(0.5)
      | 	socket_close()
      | end
      | 
      | def CW_Rotate(angle):
      | 	socket_open(SERVER_IP, SERVER_PORT)
      | 	socket_send_string("CWROTATE:"+to_str(angle))
      | 	sync()
      | 	sleep(0.5)
      | 	socket_close()
      | end
      | 
      | def CCW_Rotate(angle):
      | 	socket_open(SERVER_IP, SERVER_PORT)
      | 	socket_send_string("CCWROTATE:"+to_str(angle))
      | 	sync()
      | 	sleep(0.5)
      | 	socket_close()
      | end
      | 
      | def CW_full_Rotate():
      | 	socket_open(SERVER_IP, SERVER_PORT)
      | 	socket_send_string("FULLROTATE:"+to_str(1))
      | 	sync()
      | 	sleep(0.5)
      | 	socket_close()
      | end
      | 
      | def CCW_full_Rotate():
      | 	socket_open(SERVER_IP, SERVER_PORT)
      | 	socket_send_string("FULLROTATE:"+to_str(-1))
      | 	sync()
      | 	sleep(0.5)
      | 	socket_close()
      | end
      | 
      | def tilt_to_home():
      | 	socket_open(SERVER_IP, SERVER_PORT)
      | 	socket_send_string("HOME")
      | 	sync()
      | 	sleep(0.5)
      | 	socket_close()
      | end
      | #######
      | def vibration_1():
      | 	set_analog_out(0,0.4)
      | 	sleep(1)
      | 	set_analog_out(0,0.0)
      | 	sleep(0)
      | end
      | 
      | def vibration_2():
      | 	set_analog_out(0,0.4)
      | 	sleep(0.8)
      | 	set_analog_out(0,0.0)
      | 	sleep(0.2)
      | end
      | 
      | def vibration_3():
      | 	set_analog_out(0,0.4)
      | 	sleep(0.5)
      | 	set_analog_out(0,0.0)
      | 	sleep(0.3)
      | end
      | 
      | def vibration_4():
      | 	set_analog_out(0,0.4)
      | 	sleep(0.5)
      | 	set_analog_out(0, 0.0)
      | 	sleep(0.5)
      | end
      | 
      | def vibration_5():
      | 	set_analog_out(0,0.4)
      | 	sleep(0.2)
      | 	set_analog_out(0, 0.0)
      | 	sleep(0.8)
      | end
      | 
      | ##################
      | 
      | global gear_2_holder = 0.018
      | global gain_per_percent = 0.5
      | global w_dosed_total = 0.0
      | global last_scale = 0.0
      | global tilt_angle_sent = 0.0
      | global level = 0.0
      | global target_g = 0.0
      | global angle_max = 60
      | global angle_min = 10
      | global hinge_2_base = 0.0421
      | global TCP_2_tip_x = 0.0047
      | global spatula_len = 0.182
      | global spatula_offset = p[TCP_2_tip_x,0,spatula_len,0,0,0]
      | global SPATULA_L_VOL_ML = 5.0        # 1 teaspoon = 5 mL
      | global SPATULA_M_VOL_ML = 1.25       # 1/4 teaspoon = 1.25 mL
      | global SPATULA_S_VOL_ML = 0.15625    # 1/32 teaspoon = 0.15625 mL
      | global SPATULA_FLAT_M_VOL_ML  = 2.2
      | global SPATULA_FLAT_S_VOL_ML  = 1.2   #based on caluclations using rho = m/V
      | global ry_deg_safe = 0
      | global ry_deg = 0
      | global g_prev_cum_w = -1.0
      | global g_depth_corr = 0.0
      | global scoop_ct = 0
      | global error_sum = 0.0
      | global error_sq_sum = 0.0
      | global scoop_g = 0.0
      | #global w_dosed_total = 0.0
      | global g_corr_max = 0.01
      | global g_k = 0.0
      | global prev_weight = -1.0
      | global rep_weight = -2.0
      | 
      | def clamp(x, lo, hi):
      | 	if(x<lo):
      | 		return lo
      | 	elif (x>hi):
      | 		return hi
      | 	else:
      | 		return x
      | 	end
      | end
      | 
      | def compute_level_percent(W_now, weight_value):   # W_now = container+powder, weight_value = live scale reading
      |     global delta = weight_value - last_scale
      | 
      |     if (delta < 0.0):
      |         delta = 0.0
      |     end
      | 
      |     global w_dosed_total = w_dosed_total + delta
      |     global last_scale = weight_value     # update the last scale reading
      | 
      |     local W_eff = W_now - w_dosed_total
      |     if (W_eff <  empty_weight_g):
      |         W_eff =  empty_weight_g
      |     end
      | 
      |     # Compute powder level %
      |     level = 100.0 * (W_eff -  empty_weight_g) / (full_weight_g -  empty_weight_g)
      | 
      |     # Clamp to 0–100
      |     level = clamp(level, 0, 100)
      |   textmsg("deb 1 = ", level)
      |     return level
      | end
      | 
      | def deg2rad(d):
      | 	return d*3.141592/180
      | end
      | 
      | def my_abs(val):
      | 	if (val<0):
      | 		return -val
      | 	else:
      | 		return val
      | 	end
      | end
      | 
      | def compute_tilt_deg(level_percent):
      | 	angle = angle_min + gain_per_percent*(100.0-level_percent)
      | 
      |   	textmsg("deb 2 = ", angle)
      | 	return clamp(angle, angle_min, angle_max)
      | end
      | 
      | def tilt(level_percentage):
      | 	new_angle = compute_tilt_deg(level_percentage)
      |   	textmsg("deb angle 1 = ", new_angle)
      | 	global angle_rel = new_angle - tilt_angle_sent
      |   	textmsg("deb 2 = ", angle_rel)
      | 
      | 	if my_abs(angle_rel)>2.0:
      |   		textmsg("deb loop")
      | 		tilt_send(new_angle)
      | 		global angle_deg = new_angle
      |   		textmsg("deb 2 = ", angle_deg)
      | 		global tilt_angle_sent = new_angle
      | 		global p_center_vertical = center_pose()
      | 		global p_center = updated_center_pose(p_center_vertical, angle_deg)
      | 	end
      |   	textmsg("deb loop exit")
      | 
      | 	tilt_send(angle_deg)
      |   	textmsg("deb angle 2 =", angle_deg)
      | 
      | end
      | 
      | def compute_scoop_depth(level, weight_value, target_g):
      | 
      | 	global scoop_depth_rel = ((100.0-level)/100.0)*(H -mouth_sh)
      | 	if (g_prev_cum_w<0):
      | 		g_prev_cum_w = weight_value
      | 		g_depth_corr = 0.0
      | 	else:
      | 		global scoop_g = weight_value-g_prev_cum_w
      | 		g_prev_cum_w = weight_value
      | 
      | 		e = target_g-scoop_g
      | 
      | 		corr_proposed = g_k*e
      | 		#g_depth_corr = (1.0 -g_alpha)*g_depth_corr + g_alpha*corr_proposed
      | 		g_depth_corr = clamp(corr_proposed, -g_corr_max, g_corr_max)
      | 	end
      | 
      | 	global scoop_depth = scoop_depth_rel + g_depth_corr
      | 	global scoop_depth = clamp(scoop_depth, 0, H)
      | 	return scoop_depth
      | end
      | 
      | def get_scoop_weight(spatula, bulk_density):
      | 
      | 	local vol = 0
      | 
      | 	if (spatula == "spatula_L"):
      | 		vol = SPATULA_L_VOL_ML
      | 		global spatula_depth = 0.015
      | 		global spatula_mid   = 0.016
      | 		global spatula_ry    = 0.0
      | 
      | 	elif (spatula == "spatula_M"):
      | 		vol = SPATULA_M_VOL_ML
      | 		global spatula_depth = 0.010
      | 		global spatula_mid   = 0.0105
      | 		global spatula_ry    = 0.0
      | 
      | 	elif (spatula == "spatula_S"):
      | 		vol = SPATULA_S_VOL_ML
      | 		global spatula_depth = 0.008
      | 		global spatula_mid   = 0.0063
      | 		global spatula_ry    = 0.0
      | 
      | 	elif (spatula == "spatula_flat_M"):
      | 		vol = SPATULA_FLAT_M_VOL_ML
      | 		global spatula_depth = 0.01
      | 		global spatula_mid   = 0.02
      | 		global spatula_ry    = 7.0
      | 
      | 	elif (spatula == "spatula_flat_S"):
      | 		vol = SPATULA_FLAT_S_VOL_ML
      | 		global spatula_depth = 0.005
      | 		global spatula_mid   = 0.016
      | 		global spatula_ry    = 2.0
      | 
      | 	else:
      | 		textmsg("Unknown spatula type")
      | 		return 0.0
      | 	end
      | 	global target_g = vol * bulk_density
      | 	return target_g
      | 
      | end
      | 
      | def select_spatula(Flowability, level, diff, bulk_density, mouth_d ):
      | 
      |     local k = 1.1
      | 
      |     global powder_height = (H  - mouth_sh ) * level/100
      | 
      |     if (Flowability == "LOW"):
      | 
      |         local gFM = get_scoop_weight("spatula_flat_M", bulk_density)
      | 
      |         local level_ok_FM = (spatula_mid  < powder_height)
      |         local diff_ok_FM  = (diff > k * gFM)
      | 
      |         local flatM_ok = level_ok_FM and diff_ok_FM
      | 
      |         if (flatM_ok):
      |             return "spatula_flat_M"
      |         else:
      |             return "spatula_flat_S"
      |         end
      | 
      |     end
      | 
      |     local gL = get_scoop_weight("spatula_L", bulk_density)
      | 
      |     local mouth_ok_L = (mouth_d  >= 0.05)
      |     local level_ok_L = (spatula_mid < powder_height)
      |     local diff_ok_L  = (diff > k * gL)
      | 
      |     local large_ok = mouth_ok_L and level_ok_L and diff_ok_L
      | 
      |     local gM = get_scoop_weight("spatula_M", bulk_density)
      | 
      |     local level_ok_M = (spatula_mid < powder_height)
      |     local diff_ok_M  = (diff > k * gM)
      | 
      |     local medium_ok = level_ok_M and diff_ok_M
      | 
      |     if (large_ok):
      |         return "spatula_L"
      | 
      |     elif (medium_ok):
      |         return "spatula_M"
      | 
      |     else:
      |         return "spatula_S"
      |     end
      | 
      | end
      | 
      | def after_scoop():
      | 	set_tcp(tcp_dosing)
      | 	set_analog_out(0,0.0)
      | 	tilt_send(angle_deg)
      | 	sleep(0.5)
      | 	movel(lifted_pose, a=0.05, v=0.2)
      | 	movel(tilted_pose_in_base2, a=0.05, v=0.2)
      | 	set_analog_out(0,0.4)
      | 	movel(pose_trans(tilted_pose_in_base2, p[0,0,0,0,0,2.0]), a=0.05, v=0.2)
      | 	set_analog_out(0,0.0)
      | 	movel(tilted_pose_in_base2, a=0.05, v=0.2)
      | 	movel(lifted_pose, a=0.05, v=0.2)
      | 	tilt_to_home()
      | 	set_tcp(tcp_default)
      | end
      | 
      | def center_pose():
      | 	global p_translated = container_place
      | 	#global p_translated = pots_axis_temp
      | 
      | 	#cx = p_translated[0]
      | 	#cy = p_translated[1]
      | 	#cz = p_translated[2]
      | 
      | 	global p_center_vertical_temp = pose_trans(p_translated, p[0,0,0, deg2rad(90), 0, 0])
      | 	cx = p_center_vertical_temp[0]
      | 	cy = p_center_vertical_temp[1]
      | 	cz = p_center_vertical_temp[2]
      | 	rx = p_center_vertical_temp[3]
      | 	ry = p_center_vertical_temp[4]
      | 	rz = p_center_vertical_temp[5]
      | 
      | 	global p_center_vertical_temp = p[cx,cy,cz, 0, 0, rz]
      | 	trans_rel = p[0,0,-pick_2_base+H,0,0,0]
      | 	global p_center_vertical =  pose_trans(p_center_vertical_temp, trans_rel)
      | 	return p_center_vertical
      | end
      | 
      | def updated_center_pose(p_center_vertical, angle_deg):
      | 	hinge_pose = pose_trans(p_center_vertical, p[0,0,-hinge_2_base-gear_2_holder-H ,0,0,0])
      | 	local_rel = pose_trans(pose_inv(hinge_pose), p_center_vertical)
      | 
      | 	rot_tilt = p[0,0,0, -deg2rad(angle_deg),0,0]
      | 	local_rel_tilted = pose_trans(rot_tilt, local_rel)
      | 
      | 	global p_center = pose_trans(hinge_pose, local_rel_tilted)
      | 	return p_center
      | end
      | 
      | def scoop_powder(p_center):
      | 	vibration_voltage = 0.4
      | 	global scoop_radius_default = 0.0
      | 
      | 
      | 	scoop_radius_default = mouth_d /2 - spatula_depth
      | 	scoop_safe_entry_pose = pose_trans(p_center, p[-TCP_2_tip_x,0,spatula_len+0.05,0,0,0])
      | 	scoop_entry_pose = pose_trans(p_center, p[-TCP_2_tip_x,0,spatula_len,0,0,0])
      | 
      | 	movel(scoop_safe_entry_pose, a=0.1, v=0.25)
      | 	movel(scoop_entry_pose, a=0.1, v=0.25)
      | 
      | 	scoop_start_rel_int = p[0, 0, -mouth_sh , 0, 0, 0]
      | 	scoop_start_pose_int = pose_trans(scoop_entry_pose, scoop_start_rel_int)
      | 
      | 	movel(scoop_start_pose_int, a=0.1, v=0.25)
      | 
      | 	#local ry_deg = map_tilt_to_ry_deg(angle_deg,level)
      | 	#local ry_result = map_tilt_to_ry_deg(angle_deg,level)
      | 
      | 	#global scoop_depth = compute_scoop_depth(level,weight_value, target_g)
      | 	safe_scoop_pivot = (mouth_d  - spatula_depth)/(scoop_depth+mouth_sh+spatula_mid)
      | 	global ry_safe = asin(safe_scoop_pivot)
      | 	global ry = deg2rad(90-angle_deg)
      | 
      | 	#global ry_safe = ry_result[0]
      | 	#global ry = deg2rad(ry_result[1])
      | 
      | 	if (spatula_mid < powder_height):
      | 		global scoop_status= "normal"
      | 		global total_depth = mouth_sh + scoop_depth + spatula_mid
      | 		global total_depth = clamp(total_depth, 0, H - spatula_mid)
      | 		scoop_start_rel = p[scoop_radius_default, 0, -total_depth, 0, 0, 0]
      | 
      | 		rot_mid = p[0, 0, 0, 0, 0, 0.785]
      | 		rot_end = p[0, 0, 0, 0, 0, 1.5708]
      | 
      | 		scoop_via_rel = pose_trans(rot_mid, scoop_start_rel)
      | 		scoop_end_rel = pose_trans(rot_end, scoop_start_rel)
      | 
      | 		scoop_start_pose = pose_trans(scoop_entry_pose, scoop_start_rel)
      | 		scoop_via_pose = pose_trans(scoop_entry_pose, scoop_via_rel)
      | 		scoop_end_pose = pose_trans(scoop_entry_pose, scoop_end_rel)
      | 
      | 		movel(scoop_start_pose, a=0.1, v=0.25)
      | 
      | 		if (level<90.0):
      | 			CW_full_Rotate()
      | 		end
      | 
      | 		movec(scoop_via_pose, scoop_end_pose, a=0.03, v=0.02)
      | 		sleep(1.0)
      | 
      | 
      | 		# safe_retention
      | 		local pivot_pose = pose_trans(scoop_end_pose, p[0,0,total_depth-spatula_len,0,0,0])
      | 		local end_rel = pose_trans(pose_inv(pivot_pose), scoop_end_pose)
      | 		local end_rel_tilted = pose_trans(end_rel, p[0, 0, 0, 0, ry_safe-deg2rad(spatula_ry), 0])
      | 		local tilted_pose_in_base = pose_trans(pivot_pose, p[0,0,0,end_rel_tilted[3],end_rel_tilted[4], end_rel_tilted[5]])
      | 		local tilted_pose_in_base = pose_trans(tilted_pose_in_base, p[0, 0, spatula_len-total_depth, 0, 0, 0])
      | 		# sptula pivoted around the container rim of the mouth at ry_safe
      | 		movel(tilted_pose_in_base, a=0.03, v=0.1)
      | 
      | 		global safe_x = sin(ry_safe)*(scoop_depth - (mouth_d -spatula_depth)/tan(90-ry_safe/2))
      | 		global safe_z = cos(ry_safe)*(scoop_depth - (mouth_d -spatula_depth)/tan(90-ry_safe/2))
      | 
      | 		local safe_up = pose_trans(tilted_pose_in_base, p[-safe_x,0,safe_z,0,0,0])
      | 		movel(safe_up, a=0.03, v=0.1)
      | 
      | 		# full exit
      | 		#local pivot_pose2 = pose_trans(tilted_pose_in_base, p[0,0,total_depth-spatula_len,0,0,0])
      | 		local pivot_pose2 = pose_trans(scoop_entry_pose, p[0,0,-spatula_len,0,0,0])
      | 		local end_rel2 = pose_trans(pose_inv(pivot_pose2), tilted_pose_in_base)
      | 		#popup("is the spatula crashing front? ", blocking = True)
      | 		local end_rel_tilted2 = pose_trans(end_rel2, p[0, 0, 0, 0, ry-ry_safe-deg2rad(spatula_ry), 0])
      | 
      | 	else : # emptying logic
      | 		CCW_full_Rotate()
      | 		global scoop_status= "emptying"
      | 		spatula_base = pose_trans(scoop_entry_pose, p[0, 0, -H+wall_thickness, 0, 0, 0])
      | 		local pivot_pose2 = pose_trans(scoop_entry_pose, p[0,0,-spatula_len,0,0,0])
      | 		# tilt inwards
      | 		global in_angle = -atan((cent_edge-2*spatula_depth)/(2*H))
      | 		spatula_tilt_rel = pose_trans(pose_inv(pivot_pose2), spatula_base)
      | 
      | 		spatula_tilt = pose_trans(spatula_tilt_rel, p[0, 0, 0, -in_angle, 0, 0])
      | 		global tilted_pose = pose_trans(pivot_pose2, p[0,0,0,spatula_tilt[3],spatula_tilt[4], spatula_tilt[5]])
      | 
      | 		global tilted_pose = pose_trans(tilted_pose, p[0,0,spatula_len-H+wall_thickness,0,0,0])
      | 
      | 		movel(tilted_pose,a=0.1, v=0.25)
      | 
      | 		rotate90=pose_trans(tilted_pose,p[0,0,0,0,0,1.5708])
      | 
      | 		#sleep(1)
      | 		#Rotate()
      | 		#sleep(0.2)
      | 		movel(rotate90, a=0.1, v=0.1)
      | 		#popup("is the spatula crashing front? ", blocking = True)
      | 		movel(pose_trans(scoop_start_pose_int,p[0,0,0,0,0,1.5708]), a=0.03, v=0.1)
      | 		# full exit
      | 		#local pivot_pose2 = pose_trans(scoop_entry_pose, p[0,0,-spatula_len,0,0,0])
      | 		local end_rel2 = pose_trans(pose_inv(scoop_entry_pose), rotate90)
      | 		local end_rel_tilted2 = pose_trans(end_rel2, p[0, 0, 0, 0, ry-in_angle-deg2rad(spatula_ry), 0])
      | 	end
      | 
      | 	# exit flat spoon
      | 	global tilted_pose_in_base2 = pose_trans(pivot_pose2, p[0,0,0,end_rel_tilted2[3],end_rel_tilted2[4], end_rel_tilted2[5]])
      | 	global tilted_pose_in_base2 = pose_trans(tilted_pose_in_base2, p[0, 0, spatula_len-spatula_mid, 0, 0, 0])
      | 	# spaula exited at center of the mouth at ry
      | 	movel(tilted_pose_in_base2, a=0.03, v=0.1)
      | 	#popup("is the spatula crashing at mouth? ", blocking = True)
      | 	if(scoop_status== "normal"):
      | 
      | 		if (spatula=="spatula_flat_S" or spatula=="spatula_S"):
      | 			vibration_1()
      | 			sleep(1)
      | 			#vib_thread = False
      | 			local ry_level = deg2rad(10)
      | 		elif (spatula == "spatula_M"):
      | 			vib_thread=True
      | 			set_analog_out(0,0.4)
      | 			#vibration_3()
      | 			local ry_level = deg2rad(25)
      | 		else:
      | 			vib_thread=True
      | 			vibration_3()
      | 			local ry_level = deg2rad(10)
      | 		end
      | 
      | 		# remove excess
      | 		local pivot_pose_level = pose_trans(tilted_pose_in_base2, p[0,0,-spatula_len,0,0,0])
      | 		local end_rel_level = pose_trans(pose_inv(pivot_pose_level), tilted_pose_in_base2)
      | 		#local ry_level = ry/1.5
      | 		#local ry_level = deg2rad(15)
      | 		local end_rel_tilted_level = pose_trans(end_rel_level, p[0, 0, 0, 0, -ry_level, 0])
      | 		local end_rel_tilted_level2 = pose_trans(pivot_pose_level, p[0, 0, 0,end_rel_tilted_level[3],end_rel_tilted_level[4], end_rel_tilted_level[5]])
      | 		local end_rel_tilted_level2 = pose_trans(end_rel_tilted_level2, p[0,0,spatula_len,0,0,0])
      | 		movel(end_rel_tilted_level2, a=0.03, v=0.1)
      | 
      | 		movel(tilted_pose_in_base2, a=0.03, v=0.1)
      | 		vib_thread=False
      | 		set_analog_out(0, 0.0)
      | 	else:
      | 		set_analog_out(0, 0.0)
      | 	end
      | 	#popup("safe out + moving towards beaker", title = "Pause", blocking = True)
      | 	global lifted_pose = pose_trans(tilted_pose_in_base2, p[-0.04,0,0.04,0,0,0]) # safety distance away from the container
      | 
      | 	movel(lifted_pose, a=0.03, v=0.1)
      | 	tilt_to_home()
      | end
      | 
      | def auto_tilt_and_scoop(W_now, target_weight, weight_value):
      | 	set_tcp(tcp_dosing)
      | 	global level = compute_level_percent(W_now, weight_value)
      | 
      | 	global spatula = select_spatula(Flowability, level, diff, bulk_density, mouth_d )
      | 	textmsg("deb 4 = ", spatula)
      | 	global target_g = get_scoop_weight(spatula, bulk_density)
      | 	textmsg("deb 5 = ", target_g)
      | 	global scoop_depth = compute_scoop_depth(level, weight_value, target_g)
      |   	textmsg("deb 6 = ", scoop_depth)
      | 	tilt(level)
      | 	if (scoop_ct < 5 and g_prev_cum_w>0.0):
      | 		#local scoop_g = scoop_g
      | 		local error = target_g - scoop_g
      | 		error_sum = error_sum + error
      | 		error_sq_sum = error_sq_sum + error*error
      | 		scoop_ct = scoop_ct+1
      | 
      | 		if (scoop_ct==5):
      | 			local avg_error = error_sum/5.0
      | 			#local std_dev = sqrt(error_sq_sum/5.0) - (avg_error*avg_error)
      | 
      | 			if (my_abs(avg_error)>1.0):
      | 				global g_k = 0.055
      | 				#g_alpha = 0.85
      | 			elif (my_abs(avg_error)>0.6):
      | 				global g_k= 0.045
      | 				#g_alpha =0.75
      | 			elif (my_abs(avg_error)> 0.3):
      | 				global g_k = 0.035
      | 				#g_alpha = 0.65
      | 			elif (my_abs(avg_error)>0.1):
      | 				global g_k = 0.025
      | 				#g_alpha = 0.55
      | 			else:
      | 				global g_k = 0.015
      | 				#g_alpha = 0.45
      | 			end
      | 			global g_alpha = 0.6
      | 		end
      | 	end
      | 	scoop_powder(p_center)
      | 	#textmsg("deb 7 - sucess")
      |  	set_tcp(tcp_default)
      | end
    Script file /programs/04 Scripts/Weight_scale_socket_s.script
      | global s_depth = 0
      | global s_length =0
      | global s_volume = 0
      | global ry_theta  = 0
      | 
      | def get_weight():
      | 	socket_open(SERVER_IP,SERVER_PORT)
      | 	sleep(0.2)
      | 	textmsg("socket opened successfully!")
      | 	socket_send_string("GET_WEIGHT")
      | 	sleep(0.2)
      | 	sync()
      | 	sleep(0.2)
      | 	receiveFromServ = socket_read_ascii_float(6)
      | 	sleep(1)
      | 	#while (receiveFromServ[0] <1):
      | 		#receiveFromServ = socket_read_ascii_float(1)
      | 		#sleep(1)
      | 		#textmsg("retrying read:", receiveFromServ)
      | 	#end
      | 	textmsg("Received weight:", receiveFromServ[1])
      | 	sleep(0.2)
      | 	socket_close()
      | 	sleep(0.2)
      | 	return receiveFromServ[1]
      | end
      | 
      | def tare_scale():
      | 	socket_open(SERVER_IP,SERVER_PORT)
      | 	socket_send_string("TARE")
      | 	sleep(2)
      | 	socket_close()
      | end
      | 
      | def zero_scale():
      | 	socket_open(SERVER_IP,SERVER_PORT)
      | 	socket_send_string("ZERO")
      | 	sleep(0.5)
      | 	socket_close()
      | end
      | 
      | def log_weight():
      | 	socket_open(SERVER_IP,SERVER_PORT)
      | 	socket_send_string("LOG_WEIGHT")
      | 	sleep(0.5)
      | 	socket_close()
      | end
      | 
      | def send_target_info():
      | 	socket_open(SERVER_IP,SERVER_PORT)
      | 	socket_send_string("SET_TARGET:" + to_str(target_weight))
      | 	sleep(0.2)
      | 	socket_close()
      | end
      | def send_powder_info():
      | 	socket_open(SERVER_IP,SERVER_PORT)
      | 	socket_send_string("SET_POWDER:" + Pow_name)
      | 	sleep(0.2)
      | 	socket_close()
      | end
      | def send_spatula_info():
      | 	socket_open(SERVER_IP,SERVER_PORT)
      | 	socket_send_string("SET_SPATULA:" + spatula)
      | 	#sleep(1)
      | 
      | 	#local fl = socket_read_ascii_float(4)
      | 
      |   	#global s_depth = fl[1]
      |   	#global s_length = fl[2]
      |  	#global s_volume = fl[3]
      |  	#global ry_theta  = fl[4]
      | 	sleep(0.2)
      | 	socket_close()
      | end
      | 
      | def send_level_info():
      | 	socket_open(SERVER_IP,SERVER_PORT)
      | 	socket_send_string("SET_LEVEL:" + to_str(level))
      | 	sleep(0.2)
      | 	socket_close()
      | end
      | 
      | def get_cont_weight():
      |   socket_open(SERVER_IP, SERVER_PORT)
      |   #rq_open_and_wait()
      |   cmd = "GET_CONT_WEIGHT"
      |   socket_send_string(cmd)
      |   sync()
      |   sleep(0.5)
      |   receiveFromSer = socket_read_ascii_float(1)
      |   socket_close()
      |   return receiveFromSer[1]
      | end
  Folder BeforeStarts
    Folder uLM
      CMD_Stop := False
      CMD_Abort := False
      CMD_Clear := False
      STATE := 1
      STATE_Info := ""
      ARM_Referenced := False
      Script: zero_ftsensor()
      Folder poses init
        PSE_A := p[0,0,0,0,0,0]
        PSE_A_H := p[0,0,0,0,0,0]
        PSE_R := p[0,0,0,0,0,0]
        PSE_R_H := p[0,0,0,0,0,0]
        PSE_T := p[0,0,0,0,0,0]
        PSE_T_H := p[0,0,0,0,0,0]
        PSE_C_E := p[0,0,0,0,0,0]
        PSE_C_H := p[0,0,0,0,0,0]
        PSE_C_S := p[0,0,0,0,0,0]
      Script: init_home_by_cartesian_pose(p[0,-0.400,0.300,0,0,0])
    Folder Clearing
      Script: reset_error()
      Script: reset_warning()
    Folder uGo
      SuppressedNode
        Script: ugo_init( True ,"http://192.168.12.240:10001")
      Script: ugo_init( True ,"http://192.168.12.120:10001")
      Script: ugo_update_outputs()
    Folder App
      'ADD APPLICATION SPECIFIC COMMANDS'
    Folder Tools
      OBJ_Picked := gripper_has_object()
      If OBJ_Picked
        URCap Gripper Activate (Robotiq_Grippers, Robotiq Inc.) dataModel(ResetAndActivateKey=false)
      Else 
        URCap Gripper Activate (Robotiq_Grippers, Robotiq Inc.) dataModel(ResetAndActivateKey=true)
      Script: zero_ftsensor()
      Folder EXTT
        Set DigitalOutput pin=GRP_3F_Enable; digitalValue=0
        Set DigitalOutput pin=BarcodeTrigger; digitalValue=0
        Set DigitalOutput pin=GRP_3F_Decap; digitalValue=0
        Set DigitalOutput pin=GRP_3F_Cap; digitalValue=0
        Set DigitalOutput pin=GRP_3F_Open; digitalValue=0
      PSE_T := get_tool_free_pose(dir=[0,0,0.150], move_in_base_frame=True)
      If is_reachable(Base, [PSE_T])
        MoveL speed 150 mm/s, acceleration 1200 mm/s^2 (useActiveTCP=true optimoveEnabled=false optiMoveSpeed=0.3 optiMoveAcceleration=0.09) feature=Base
          Waypoint Variable (Variable): variable=PSE_T
  Folder powder dispensing variable init
    Start_thread := False
    vib_thread := False
    w_full_thread := False
    d_cc := 0.07
    kp := 0.0035
    ki := 0.0001
    kd := 0.003
    dt := 0.2
    Integral_error := 0
    current_error := 0
    previous_error := 0
    tilt_increment := 0
    tilt_angle := 0
    diff := 0
    Script: tilt_to_home()
    Script: tilt_to_home()
    switch_spat_M := True
    switch_spat_S := True
    switch_spat_F_M := True
    switch_spat_F_S := True
    last_scale := 0
Robot Program (runOnlyOnce=false)
  Folder MAIN
    Script: command_manager(external_control="uGO", cond_suspend=(ITM_Manipulated and AMR_AtTarget and AMR_Charging and AMR_Battery<40), cond_unsuspend=(AMR_Battery≟60))
    Script: log_state(STATE_Info)
    Switch expression=STATE
      Case (caseValue=1)
        Folder Stopping [hidden by the author, left out]
      Case (caseValue=2)
        Folder Stopped [hidden by the author, left out]
      Case (caseValue=3)
        Folder  Resetting [hidden by the author, left out]
      Case (caseValue=4)
        Folder Idle [hidden by the author, left out]
      Case (caseValue=5)
        Folder Starting
          STATE_Info := "Starting"
          'ADD COMMANDS WHAT TO START WITH'
          Call Sub_AMR_MiR_V3
          Folder get ugo data
            Folder Assign Tasks
              Script: TASK.ID = ugo_get_task()
              If TASK.ID≟1
                Task_info := "Charge"
                Folder Parameters [hidden by the author, left out]
              ElseIf TASK.ID≟9
                'Pick Sarstedt Rack from Variable source'
                Task_info := "Navigate to Target"
                Folder Parameters [hidden by the author, left out]
              ElseIf TASK.ID≟13
                Task_info := "Dose Powder"
                Folder Parameters
                  ITM_ID := 1
                  W_now := (UGO.read_input("00","Container_weight"))/1000
                  Pow_name := (UGO.read_input("00","Powder_name"))
                  target_weight := (UGO.read_input("00","Target_weight"))/1000
                  Script: send_picking_info(Pow_name,target_weight)
                  w_dosed_total := 0
                  OBJ_Type := 6
                  JIG := 17
                  AMR_PosTarget := 5
              ElseIf TASK.ID≟49
                Task_info := "Pick Containers"
                Folder Parameters
                  ITM_ID := 1
                  OBJ_Type := 6
                  JIG := 15
                  AMR_PosTarget := 3
              ElseIf TASK.ID≟50
                Task_info := "Decap Containers"
                Folder Parameters
                  ITM_ID := 1
                  OBJ_Type := 6
                  JIG := 16
                  AMR_PosTarget := 5
              ElseIf TASK.ID≟51
                Task_info := "Detect Spatula and transfer powder"
                Folder Parameters
                  ITM_ID := 1
                  target_weight := (UGO.read_input("00","Target_weight"))/1000
                  OBJ_Type := 8
                  JIG := 16
                  AMR_PosTarget := 5
              ElseIf TASK.ID≟52
                Task_info := "Pick Powder"
                Folder Parameters
                  ITM_ID := 1
                  SuppressedNode
                    Pow_name := (UGO.read_input("00","Powder_name"))
                  OBJ_Type := 6
                  JIG := 15
                  AMR_PosTarget := 3
              ElseIf TASK.ID≟53
                Task_info := "Decap Powder"
                Folder Parameters
                  ITM_ID := 1
                  OBJ_Type := 6
                  JIG := 1
                  AMR_PosTarget := 5
              ElseIf TASK.ID≟54
                Task_info := "Empty and swap Powder container"
                SuppressedNode
                  Folder Parameters
                    ITM_ID := 1
                    target_weight := (UGO.read_input("00","Target_weight"))/1000
                    W_now := (UGO.read_input("00","Container_weight"))/1000
                    Pow_name := (UGO.read_input("00","Powder_name"))
                    OBJ_Type := 6
                    JIG := 17
                    AMR_PosTarget := 5
                Folder Parameters
                  ITM_ID := 1
                  SuppressedNode
                    target_weight := (UGO.read_input("00","target_weight"))/1000
                  W_now := (UGO.read_input("00","Container_weight"))/1000
                  Pow_name := (UGO.read_input("00","Powder_name"))
                  SuppressedNode
                    Script: scooping_init()
                  SuppressedNode
                    target_weight := W_now-W_EMPTY-(0.002*W_FULL)
                  OBJ_Type := 6
                  JIG := 17
                  AMR_PosTarget := 5
              ElseIf TASK.ID≟55
                Task_info := "Place Powder"
                Folder Parameters
                  ITM_ID := 1
                  OBJ_Type := 6
                  JIG := 21
                  AMR_PosTarget := 5
              ElseIf TASK.ID≟56
                Task_info := "Dose Powder"
                Folder Parameters
                  ITM_ID := 1
                  target_weight := (UGO.read_input("00","Target_weight"))/1000
                  W_now := (UGO.read_input("00","Container_weight"))/1000
                  Pow_name := (UGO.read_input("00","Powder_name"))
                  OBJ_Type := 6
                  JIG := 17
                  AMR_PosTarget := 5
              ElseIf TASK.ID≟57
                Task_info := "Recipe Powder dosing"
                Folder Parameters
                  ITM_ID := 1
                  Pow_A := (UGO.read_input("00","PowderA"))
                  Pow_B := (UGO.read_input("00","PowderB"))
                  Pow_C := (UGO.read_input("00","PowderC"))
                  Total_weight := (UGO.read_input("00","Total_weight"))/1000
                  Pow_A_percent := (UGO.read_input("00","PowderA_percentage"))/100
                  Pow_B_percent := (UGO.read_input("00","PowderB_percentage"))/100
                  Pow_C_percent := (UGO.read_input("00","PowderC_percentage"))/100
                  OBJ_Type := 6
                  JIG := 17
                  AMR_PosTarget := 5
              ElseIf TASK.ID≟58
                Task_info := "Pick Powder containers"
                Folder Parameters [hidden by the author, left out]
              ElseIf TASK.ID≟59
                Task_info := "Empty Powder container"
                Folder Parameters
                  ITM_ID := 1
                  SuppressedNode
                    W_now := (UGO.read_input("00","Container_weight"))/1000
                  Pow_name := (UGO.read_input("00","Powder_name"))
                  SuppressedNode
                    Script: global target_weight = to_str(aa_weight_cont-empty_weight_g)
                  target_weight := aa_weight_cont-empty_weight_g
                  Script: send_picking_info(Pow_name,target_weight)
                  w_dosed_total := 0
                  OBJ_Type := 6
                  JIG := 17
                  AMR_PosTarget := 5
              ElseIf TASK.ID≟61
                Task_info := "Weigh, Place & Decap"
                Folder Parameters
                  ITM_ID := 1
                  OBJ_Type := 6
                  JIG := 21
                  AMR_PosTarget := 5
              Else 
                Script: set_error(ERROR_WRONG_ORDER)
          Folder test ugo
            Wait Sleep waitTime=0.2
            Script: ugo_update_outputs()
          If starting() and AMR_Done
            Script: log_message(Task_info, "New Task: ")
            Script: log_message(to_str(TASK.ID), "Task_ID: ")
            Script: do_transition(keep_rxry=OBJ_Picked)
            STATE := 6
            Script: ugo_update_outputs()
      Case (caseValue=6)
        Folder Execute
          STATE_Info := "Execute"
          If not CMD_Hold and not CMD_Suspend (checkContinuously=true)
            Switch expression=PROCESS_Step
              Case (caseValue=0)
                PROCESS_Info := "process control"
                Script: log_process(PROCESS_Info)
                Folder process control [hidden by the author, left out]
              Case (caseValue=1)
                Folder navigate [hidden by the author, left out]
              Case (caseValue=2)
                Folder prepare [hidden by the author, left out]
              Case (caseValue=3)
                Folder work
                  'ADD EVERY MACHINE, OBJECT, STATION TO WORK ON'
                  Switch expression=ITM_ID
                    Case (caseValue=1)
                      Folder uLM
                        If TASK.ID≟12
                          Folder fill racks [hidden by the author, left out]
                        ElseIf TASK.ID≟13
                          Folder Dose Powder
                            Action := 131
                            Call Sub_Vision_V18
                            Action := 34
                            Call Sub_Action_V4
                            PROCESS_Step := 0
                            WRK_Done := True
                        ElseIf TASK.ID≟49
                          Folder Pick Powder container [hidden by the author, left out]
                        ElseIf TASK.ID≟50
                          Folder Decap containers [hidden by the author, left out]
                        ElseIf TASK.ID≟51
                          Folder Detect Spatula and transfer powder [hidden by the author, left out]
                        ElseIf TASK.ID≟52
                          Folder Pick Powder container
                            Action := 131
                            Call Sub_Vision_V18
                            Action := 39
                            Call Sub_Action_V4
                            PROCESS_Step := 0
                            WRK_Done := True
                        ElseIf TASK.ID≟53
                          Folder Decap containerA
                            Action := 40
                            Call Sub_Action_V4
                            PROCESS_Step := 0
                            WRK_Done := True
                        ElseIf TASK.ID≟55
                          Folder Place Powder
                            Action := 131
                            Call Sub_Vision_V18
                            Action := 41
                            Call Sub_Action_V4
                            PROCESS_Step := 0
                            WRK_Done := True
                        ElseIf TASK.ID≟54
                          Folder Empty and swap container
                            Action := 131
                            Call Sub_Vision_V18
                            Action := 42
                            Call Sub_Action_V4
                            PROCESS_Step := 0
                            WRK_Done := True
                        ElseIf TASK.ID≟56
                          Folder Dispense Powder [hidden by the author, left out]
                        ElseIf TASK.ID≟57
                          Folder Recipe Dosing
                            Action := 48
                            Call Sub_Action_V4
                            SuppressedNode
                              Script: recipe_init(Pow_A, Pow_B, Pow_C, Total_weight, Pow_A_percent, Pow_B_percent, Pow_C_percent)
                            SuppressedNode
                              Loop While (checkContinuously=false) expression=recipe_next()≟ True
                                Action := 44
                                Call Sub_Action_V4
                                JIG := 21
                                Action := 131
                                Call Sub_Vision_V18
                                Action := 45
                                Call Sub_Action_V4
                                Script: dosing_start()
                                JIG := 17
                                Action := 131
                                Call Sub_Vision_V18
                                Action := 46
                                Call Sub_Action_V4
                                Script: dosing_end()
                            PROCESS_Step := 0
                            WRK_Done := True
                        ElseIf TASK.ID≟58
                          Folder Pick Powder containers
                            Num_cont_picked := 0
                            powder_position := "Position1"
                            Loop While (checkContinuously=false) expression=Num_cont_picked<3
                              Action := 131
                              Call Sub_Vision_V18
                              Action := 47
                              Call Sub_Action_V4
                            PROCESS_Step := 0
                            WRK_Done := True
                        ElseIf TASK.ID≟59
                          Folder Empty powder container
                            Action := 131
                            Call Sub_Vision_V18
                            Action := 50
                            Call Sub_Action_V4
                            PROCESS_Step := 0
                            WRK_Done := True
                        ElseIf TASK.ID≟61
                          Folder Place Powder
                            Action := 131
                            Call Sub_Vision_V18
                            Action := 51
                            Call Sub_Action_V4
                            PROCESS_Step := 0
                            WRK_Done := True
                    Case (caseValue=2)
                      SuppressedNode
                        Folder Centrfiuge
                          SuppressedNode
                            Script: cent_error_check()
                          OBJ_Type := 1
                          If not ERROR.FLAG
                            'load racks'
                            If TASK.ID≟14
                              Loop While (checkContinuously=false) expression=(PRC_RackCounter<4) and  not CMD_Stop and  not ERROR.FLAG
                                ITM_ID := TASK.WORK.ITM_ID_Src
                                JIG := 4
                                JIG_Slot := PRC_RackCounter+1
                                Action := 1
                                CallSubProgram
                                If OBJ_Picked and  not ERROR.FLAG
                                  ITM_ID := TASK.WORK.ITM_ID_Tgt
                                  Script: execute_cent_action(ACTION_ROTATE, JIG_Slot)
                                  Action := 7
                                  CallSubProgram
                                  PRC_RackCounter := PRC_RackCounter + 1
                              If not ERROR.FLAG
                                WRK_Done := True
                                PROCESS_Step := 0
                            'unload racks'
                            If TASK.ID≟15
                              If CNT_State_Actual≟2 or CNT_State_Actual≟3
                                Loop While (checkContinuously=false) expression=(PRC_RackCounter<4) and  not CMD_Stop and  not ERROR.FLAG
                                  ITM_ID := TASK.WORK.ITM_ID_Src
                                  JIG_Slot := PRC_RackCounter + 1
                                  Script: execute_cent_action(ACTION_ROTATE, JIG_Slot)
                                  Script: execute_cent_action(ACTION_INSPECT, JIG_Slot)
                                  Action := 8
                                  CallSubProgram
                                  If OBJ_Picked and  not ERROR.FLAG
                                    ITM_ID := TASK.WORK.ITM_ID_Tgt
                                    JIG := 4
                                    JIG_Slot := PRC_RackCounter + 1
                                    Action := 2
                                    CallSubProgram
                                    PRC_RackCounter := PRC_RackCounter+1
                                If not ERROR.FLAG
                                  WRK_Done := True
                                  PROCESS_Step := 0
                    Case (caseValue=5)
                      SuppressedNode
                        Folder SarstedtTable
                          Action := 131
                          CallSubProgram
                          Action := 1
